ABB RAPID module: MainProgram.mod

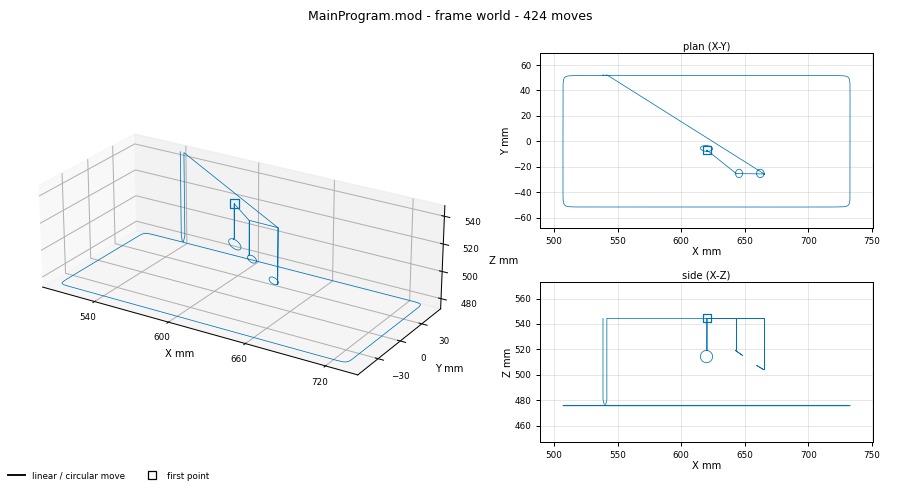
[picture p0: tool path of MainProgram.mod in frame world, 424 of 456 moves have a stored position in this frame; points joined in program order, loops and branches not executed]
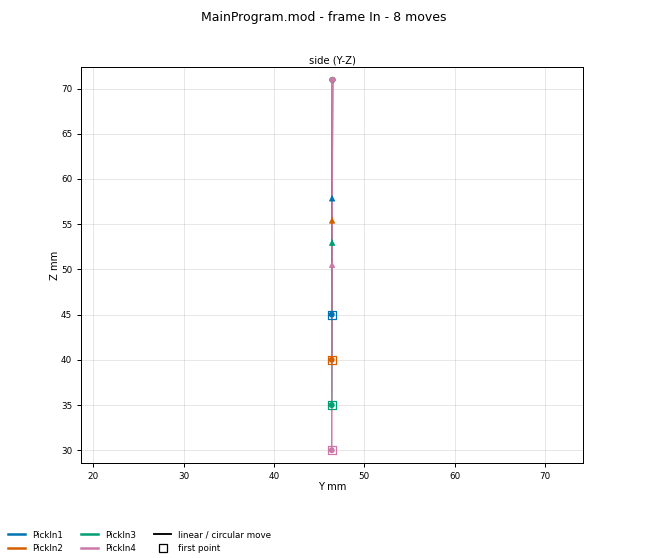
[picture p1: tool path of MainProgram.mod in frame In, 8 of 456 moves have a stored position in this frame; points joined in program order, loops and branches not executed]
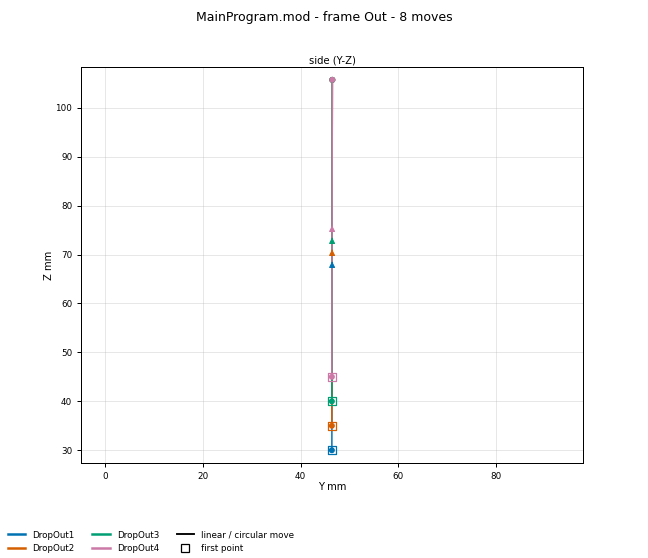
[picture p2: tool path of MainProgram.mod in frame Out, 8 of 456 moves have a stored position in this frame; points joined in program order, loops and branches not executed]
%%%
  VERSION:1
  LANGUAGE:ENGLISH
%%%
MODULE MOD_MainProgram

    ! -------------------------------
    ! Define customized variables here
    ! ...

	! Tool variables:
	PERS tooldata SuctionCup := [TRUE,[[-94.709,0.000,259.352],[0.00000000,0.00000000,0.00000000,1.00000000]],[1,[0,0,20],[1,0,0,0],0,0,0.005]];
	PERS tooldata Spindle := [TRUE,[[186.140,-0.004,258.607],[0.87136628,0.00000000,0.49063307,0.00000000]],[1,[0,0,20],[1,0,0,0],0,0,0.005]];

	! Reference variables:
	PERS wobjdata World := [FALSE, TRUE, "", [[0,0,0],[1,0,0,0]],[[390.000,0.000,0.000],[1.00000000,0.00000000,0.00000000,0.00000000]]];
	PERS wobjdata In := [FALSE, TRUE, "", [[0,0,0],[1,0,0,0]],[[290.000,450.000,10.000],[1.00000000,0.00000000,0.00000000,0.00000000]]];
	PERS wobjdata PartStation := [FALSE, TRUE, "", [[0,0,0],[1,0,0,0]],[[620.000,0.000,396.884],[0.70710678,0.00000000,0.00000000,-0.70710678]]];
	PERS wobjdata Deburring := [FALSE, TRUE, "", [[0,0,0],[1,0,0,0]],[[620.000,0.000,458.384],[0.70710678,0.00000000,0.00000000,-0.70710678]]];
	PERS wobjdata Out := [FALSE, TRUE, "", [[0,0,0],[1,0,0,0]],[[290.000,-450.000,10.000],[1.00000000,0.00000000,0.00000000,0.00000000]]];

	PROC GoHome()
		ConfJ \On;
		ConfL \Off;
		World := [FALSE, TRUE, "", [[0,0,0],[1,0,0,0]],[[390.000,0.000,0.000],[1.00000000,0.00000000,0.00000000,0.00000000]]];
		MoveAbsJ [[0.000000,0.000000,-20.000000,0.000000,30.170000,0.000000],[9E+09,9E+09,9E+09,9E+09,9E+09,9E+09]],v500,z1,SuctionCup \WObj:=World;
	ENDPROC

	PROC PickIn1()
		ConfJ \On;
		ConfL \Off;
		SuctionCup := [TRUE,[[-94.709,0.000,259.352],[0.00000000,0.00000000,0.00000000,1.00000000]],[1,[0,0,20],[1,0,0,0],0,0,0.005]];
		MoveAbsJ [[70.152800,32.938500,23.515600,0.000000,33.545900,70.152800],[9E+09,9E+09,9E+09,9E+09,9E+09,9E+09]],v500,z1,SuctionCup \WObj:=In;
		MoveL [[-16.111,46.392,45.000],[0.00000000,1.00000000,0.00000000,-0.00000000],[0,2,-2,1],[9E+09,9E+09,9E+09,9E+09,9E+09,9E+09]],v500,z1,SuctionCup \WObj:=In;
		! Attach to Suction Cup
		WaitTime 0.500;
		MoveL [[-16.087,46.472,70.960],[0.00000000,1.00000000,0.00000000,-0.00000000],[0,0,0,0],[9E+09,9E+09,9E+09,9E+09,9E+09,9E+09]],v500,z1,SuctionCup \WObj:=In;
	ENDPROC

	PROC DropStation()
		ConfJ \On;
		ConfL \Off;
		SuctionCup := [TRUE,[[-94.709,0.000,259.352],[0.00000000,0.00000000,0.00000000,1.00000000]],[1,[0,0,20],[1,0,0,0],0,0,0.005]];
		MoveAbsJ [[9.440500,34.191600,-49.511700,0.000000,105.320000,99.440500],[9E+09,9E+09,9E+09,9E+09,9E+09,9E+09]],v500,z1,SuctionCup \WObj:=PartStation;
		MoveL [[-16.111,46.392,100.500],[0.00000000,1.00000000,0.00000000,-0.00000000],[0,2,-1,1],[9E+09,9E+09,9E+09,9E+09,9E+09,9E+09]],v500,z1,SuctionCup \WObj:=PartStation;
		! Detach from Suction Cup
		WaitTime 0.500;
		MoveL [[-16.111,46.485,191.000],[0.00000000,1.00000000,0.00000000,-0.00000000],[0,0,1,0],[9E+09,9E+09,9E+09,9E+09,9E+09,9E+09]],v500,z1,SuctionCup \WObj:=PartStation;
	ENDPROC

	PROC Station1()
		ConfJ \On;
		ConfL \Off;
		! show Spindle
		TPWrite "/'Plastic deburring v9'";
		TPWrite "/''";
		TPWrite "/'NEW SECTION'";
		TPWrite "/'Strategy: swarf5d'";
		TPWrite "/'Comment: Swarf8'";
		TPWrite "/'MATRIX DEFINITION'";
		TPWrite "/'Output x(i),y(i),z(i)'";
		TPWrite "/'Output x(j),y(j),z(j)'";
		TPWrite "/'Output x(k),y(k),z(k)'";
		TPWrite "/'Output dx,dy,dz'";
		SetTool 3;
		SetRPM 5000.0;
		Spindle 1;
		MoveAbsJ [[35.301800,13.650800,12.157300,-89.295200,63.027800,42.556000],[9E+09,9E+09,9E+09,9E+09,9E+09,9E+09]],v1000,z1,Spindle \WObj:=Deburring;
		MoveL [[6.917,0.414,86.000],[0.38548738,-0.58483375,0.59278955,-0.39745378],[0,-1,0,0],[9E+09,9E+09,9E+09,9E+09,9E+09,9E+09]],v1000,z1,Spindle \WObj:=Deburring;
		MoveL [[6.917,0.414,86.000],[0.38548738,-0.58483375,0.59278955,-0.39745378],[0,-1,0,0],[9E+09,9E+09,9E+09,9E+09,9E+09,9E+09]],v1000,z1,Spindle \WObj:=Deburring;
		MoveL [[6.917,0.414,61.098],[0.38548738,-0.58483375,0.59278955,-0.39745378],[0,-2,0,0],[9E+09,9E+09,9E+09,9E+09,9E+09,9E+09]],v1000,z1,Spindle \WObj:=Deburring;
		MoveL [[7.874,0.393,60.697],[0.38548738,-0.58483375,0.59278955,-0.39745378],[0,-2,0,0],[9E+09,9E+09,9E+09,9E+09,9E+09,9E+09]],[16.67,500,5000,1000],z1,Spindle \WObj:=Deburring;
		MoveL [[7.903,0.385,60.695],[0.38548738,-0.58483375,0.59278955,-0.39745378],[0,-2,0,0],[9E+09,9E+09,9E+09,9E+09,9E+09,9E+09]],[16.67,500,5000,1000],z1,Spindle \WObj:=Deburring;
		MoveL [[7.923,0.368,60.712],[0.38548738,-0.58483375,0.59278955,-0.39745378],[0,-2,0,0],[9E+09,9E+09,9E+09,9E+09,9E+09,9E+09]],[16.67,500,5000,1000],z1,Spindle \WObj:=Deburring;
		MoveL [[7.932,0.350,60.736],[0.38548738,-0.58483375,0.59278955,-0.39745378],[0,-2,0,0],[9E+09,9E+09,9E+09,9E+09,9E+09,9E+09]],[16.67,500,5000,1000],z1,Spindle \WObj:=Deburring;
		MoveL [[7.942,0.339,60.763],[0.38548738,-0.58483375,0.59278955,-0.39745378],[0,-2,0,0],[9E+09,9E+09,9E+09,9E+09,9E+09,9E+09]],[16.67,500,5000,1000],z1,Spindle \WObj:=Deburring;
		MoveL [[7.946,0.311,60.775],[0.38548738,-0.58483375,0.59278955,-0.39745378],[0,-2,0,0],[9E+09,9E+09,9E+09,9E+09,9E+09,9E+09]],[16.67,500,5000,1000],z1,Spindle \WObj:=Deburring;
		MoveL [[7.938,0.025,60.788],[0.38288630,-0.58214828,0.59447297,-0.40137683],[0,-2,0,0],[9E+09,9E+09,9E+09,9E+09,9E+09,9E+09]],[16.67,500,5000,1000],z1,Spindle \WObj:=Deburring;
		MoveL [[7.910,-0.405,60.779],[0.38300483,-0.58012093,0.59439635,-0.40430185],[0,-2,0,0],[9E+09,9E+09,9E+09,9E+09,9E+09,9E+09]],[16.67,500,5000,1000],z1,Spindle \WObj:=Deburring;
		MoveL [[7.848,-0.934,60.707],[0.38194021,-0.57666146,0.59508111,-0.40922086],[0,-2,0,0],[9E+09,9E+09,9E+09,9E+09,9E+09,9E+09]],[16.67,500,5000,1000],z1,Spindle \WObj:=Deburring;
		MoveL [[7.772,-1.372,60.601],[0.37995322,-0.57413190,0.59635187,-0.41276211],[0,-1,0,0],[9E+09,9E+09,9E+09,9E+09,9E+09,9E+09]],[16.67,500,5000,1000],z1,Spindle \WObj:=Deburring;
		MoveL [[7.660,-1.869,60.426],[0.37743363,-0.57188089,0.59794992,-0.41587499],[0,-1,0,0],[9E+09,9E+09,9E+09,9E+09,9E+09,9E+09]],[16.67,500,5000,1000],z1,Spindle \WObj:=Deburring;
		MoveL [[7.526,-2.338,60.200],[0.37439771,-0.57017304,0.59985541,-0.41821351],[0,-1,0,0],[9E+09,9E+09,9E+09,9E+09,9E+09,9E+09]],[16.67,500,5000,1000],z1,Spindle \WObj:=Deburring;
		MoveL [[7.336,-2.857,59.865],[0.36917090,-0.56926904,0.60308585,-0.41944375],[0,-1,0,0],[9E+09,9E+09,9E+09,9E+09,9E+09,9E+09]],[16.67,500,5000,1000],z1,Spindle \WObj:=Deburring;
		MoveL [[7.162,-3.251,59.544],[0.36551673,-0.56883653,0.60530778,-0.42002978],[0,-1,0,0],[9E+09,9E+09,9E+09,9E+09,9E+09,9E+09]],[16.67,500,5000,1000],z1,Spindle \WObj:=Deburring;
		MoveL [[6.973,-3.606,59.186],[0.36224838,-0.56788024,0.60726923,-0.42132199],[0,-1,0,0],[9E+09,9E+09,9E+09,9E+09,9E+09,9E+09]],[16.67,500,5000,1000],z1,Spindle \WObj:=Deburring;
		MoveL [[6.815,-3.864,58.879],[0.36043999,-0.56727725,0.60834425,-0.42213363],[0,-1,0,0],[9E+09,9E+09,9E+09,9E+09,9E+09,9E+09]],[16.67,500,5000,1000],z1,Spindle \WObj:=Deburring;
		MoveL [[6.554,-4.204,58.361],[0.35672537,-0.56741746,0.61052971,-0.42194538],[0,-1,0,0],[9E+09,9E+09,9E+09,9E+09,9E+09,9E+09]],[16.67,500,5000,1000],z1,Spindle \WObj:=Deburring;
		MoveL [[6.282,-4.474,57.808],[0.35340770,-0.56800021,0.61245687,-0.42115952],[0,-1,0,0],[9E+09,9E+09,9E+09,9E+09,9E+09,9E+09]],[16.67,500,5000,1000],z1,Spindle \WObj:=Deburring;
		MoveL [[6.084,-4.622,57.400],[0.35045021,-0.56898176,0.61415334,-0.41983338],[0,-1,0,0],[9E+09,9E+09,9E+09,9E+09,9E+09,9E+09]],[16.67,500,5000,1000],z1,Spindle \WObj:=Deburring;
		MoveL [[5.801,-4.764,56.806],[0.34689032,-0.56972554,0.61617155,-0.41882280],[0,-1,0,0],[9E+09,9E+09,9E+09,9E+09,9E+09,9E+09]],[16.67,500,5000,1000],z1,Spindle \WObj:=Deburring;
		MoveL [[5.517,-4.832,56.200],[0.34354127,-0.57095868,0.61804469,-0.41714067],[0,-1,0,0],[9E+09,9E+09,9E+09,9E+09,9E+09,9E+09]],[16.67,500,5000,1000],z1,Spindle \WObj:=Deburring;
		MoveL [[5.234,-4.822,55.590],[0.34057760,-0.57257464,0.61968277,-0.41491981],[0,-1,0,0],[9E+09,9E+09,9E+09,9E+09,9E+09,9E+09]],[16.67,500,5000,1000],z1,Spindle \WObj:=Deburring;
		MoveL [[4.956,-4.736,54.983],[0.33797772,-0.57446132,0.62110430,-0.41230413],[0,-1,0,0],[9E+09,9E+09,9E+09,9E+09,9E+09,9E+09]],[16.67,500,5000,1000],z1,Spindle \WObj:=Deburring;
		MoveL [[4.687,-4.572,54.389],[0.33604086,-0.57652798,0.62215522,-0.40940801],[0,-1,0,0],[9E+09,9E+09,9E+09,9E+09,9E+09,9E+09]],[16.67,500,5000,1000],z1,Spindle \WObj:=Deburring;
		MoveL [[4.440,-4.339,53.840],[0.33425295,-0.57979674,0.62311733,-0.40476598],[0,-1,0,0],[9E+09,9E+09,9E+09,9E+09,9E+09,9E+09]],[16.67,500,5000,1000],z1,Spindle \WObj:=Deburring;
		MoveL [[4.245,-4.095,53.402],[0.33283353,-0.58190363,0.62387648,-0.40173143],[0,-1,0,0],[9E+09,9E+09,9E+09,9E+09,9E+09,9E+09]],[16.67,500,5000,1000],z1,Spindle \WObj:=Deburring;
		MoveL [[4.097,-3.868,53.067],[0.33181431,-0.58289839,0.62441871,-0.40028740],[0,-1,0,0],[9E+09,9E+09,9E+09,9E+09,9E+09,9E+09]],[16.67,500,5000,1000],z1,Spindle \WObj:=Deburring;
		MoveL [[3.907,-3.500,52.631],[0.32892812,-0.58510481,0.62594413,-0.39705490],[0,-1,0,0],[9E+09,9E+09,9E+09,9E+09,9E+09,9E+09]],[16.67,500,5000,1000],z1,Spindle \WObj:=Deburring;
		MoveL [[3.755,-3.123,52.278],[0.32712779,-0.58752921,0.62688678,-0.39345876],[0,-1,0,0],[9E+09,9E+09,9E+09,9E+09,9E+09,9E+09]],[16.67,500,5000,1000],z1,Spindle \WObj:=Deburring;
		MoveL [[3.623,-2.706,51.964],[0.32579005,-0.59003824,0.62758358,-0.38968521],[0,-1,0,0],[9E+09,9E+09,9E+09,9E+09,9E+09,9E+09]],[16.67,500,5000,1000],z1,Spindle \WObj:=Deburring;
		MoveL [[3.513,-2.253,51.695],[0.32545472,-0.59261817,0.62775754,-0.38575044],[0,-1,0,0],[9E+09,9E+09,9E+09,9E+09,9E+09,9E+09]],[16.67,500,5000,1000],z1,Spindle \WObj:=Deburring;
		MoveL [[3.426,-1.769,51.476],[0.32546867,-0.59528891,0.62774999,-0.38161657],[0,-1,0,0],[9E+09,9E+09,9E+09,9E+09,9E+09,9E+09]],[16.67,500,5000,1000],z1,Spindle \WObj:=Deburring;
		MoveL [[3.367,-1.261,51.311],[0.32642133,-0.59790109,0.62725498,-0.37751104],[0,-1,0,0],[9E+09,9E+09,9E+09,9E+09,9E+09,9E+09]],[16.67,500,5000,1000],z1,Spindle \WObj:=Deburring;
		MoveL [[3.336,-0.734,51.202],[0.32721447,-0.60077200,0.62684183,-0.37292496],[0,-1,0,0],[9E+09,9E+09,9E+09,9E+09,9E+09,9E+09]],[16.67,500,5000,1000],z1,Spindle \WObj:=Deburring;
		MoveL [[3.334,-0.198,51.154],[0.32817251,-0.60371090,0.62634061,-0.36814859],[0,-1,0,0],[9E+09,9E+09,9E+09,9E+09,9E+09,9E+09]],[16.67,500,5000,1000],z1,Spindle \WObj:=Deburring;
		MoveL [[3.362,0.339,51.167],[0.32965343,-0.60642410,0.62556274,-0.36366150],[0,-1,0,0],[9E+09,9E+09,9E+09,9E+09,9E+09,9E+09]],[16.67,500,5000,1000],z1,Spindle \WObj:=Deburring;
		MoveL [[3.419,0.869,51.239],[0.33178536,-0.60854381,0.62443456,-0.36010330],[0,-1,0,0],[9E+09,9E+09,9E+09,9E+09,9E+09,9E+09]],[16.67,500,5000,1000],z1,Spindle \WObj:=Deburring;
		MoveL [[3.511,1.417,51.385],[0.33673317,-0.61021010,0.62178053,-0.35727213],[0,-1,0,0],[9E+09,9E+09,9E+09,9E+09,9E+09,9E+09]],[16.67,500,5000,1000],z1,Spindle \WObj:=Deburring;
		MoveL [[3.596,1.815,51.527],[0.33843795,-0.61063438,0.62085393,-0.35654705],[0,-1,0,0],[9E+09,9E+09,9E+09,9E+09,9E+09,9E+09]],[16.67,500,5000,1000],z1,Spindle \WObj:=Deburring;
		MoveL [[3.725,2.284,51.756],[0.34227325,-0.61131950,0.61874797,-0.35537084],[0,-1,0,0],[9E+09,9E+09,9E+09,9E+09,9E+09,9E+09]],[16.67,500,5000,1000],z1,Spindle \WObj:=Deburring;
		MoveL [[3.876,2.722,52.031],[0.34580120,-0.61257678,0.61678310,-0.35319942],[0,-1,0,0],[9E+09,9E+09,9E+09,9E+09,9E+09,9E+09]],[16.67,500,5000,1000],z1,Spindle \WObj:=Deburring;
		MoveL [[4.045,3.123,52.347],[0.34927682,-0.61344264,0.61482152,-0.35169353],[0,-1,0,0],[9E+09,9E+09,9E+09,9E+09,9E+09,9E+09]],[16.67,500,5000,1000],z1,Spindle \WObj:=Deburring;
		MoveL [[4.270,3.549,52.777],[0.35456914,-0.61410907,0.61178476,-0.35052844],[0,-1,0,0],[9E+09,9E+09,9E+09,9E+09,9E+09,9E+09]],[16.67,500,5000,1000],z1,Spindle \WObj:=Deburring;
		MoveL [[4.470,3.860,53.168],[0.35787236,-0.61441666,0.60985864,-0.34998855],[0,-1,0,0],[9E+09,9E+09,9E+09,9E+09,9E+09,9E+09]],[16.67,500,5000,1000],z1,Spindle \WObj:=Deburring;
		MoveL [[4.682,4.127,53.589],[0.36134434,-0.61410206,0.60780784,-0.35054039],[0,-1,0,0],[9E+09,9E+09,9E+09,9E+09,9E+09,9E+09]],[16.67,500,5000,1000],z1,Spindle \WObj:=Deburring;
		MoveL [[4.909,4.360,54.045],[0.36290006,-0.61402146,0.60688026,-0.35068155],[0,-1,0,0],[9E+09,9E+09,9E+09,9E+09,9E+09,9E+09]],[16.67,500,5000,1000],z1,Spindle \WObj:=Deburring;
		MoveL [[5.207,4.574,54.652],[0.36756237,-0.61295146,0.60406786,-0.35254849],[0,-2,0,0],[9E+09,9E+09,9E+09,9E+09,9E+09,9E+09]],[16.67,500,5000,1000],z1,Spindle \WObj:=Deburring;
		MoveL [[5.440,4.682,55.130],[0.37069589,-0.61194017,0.60215000,-0.35430095],[0,-2,0,0],[9E+09,9E+09,9E+09,9E+09,9E+09,9E+09]],[16.67,500,5000,1000],z1,Spindle \WObj:=Deburring;
		MoveL [[5.682,4.750,55.631],[0.37301034,-0.61212853,0.60071915,-0.35397521],[0,-2,0,0],[9E+09,9E+09,9E+09,9E+09,9E+09,9E+09]],[16.67,500,5000,1000],z1,Spindle \WObj:=Deburring;
		MoveL [[5.972,4.756,56.238],[0.37688431,-0.61142117,0.59829589,-0.35519628],[0,-2,0,0],[9E+09,9E+09,9E+09,9E+09,9E+09,9E+09]],[16.67,500,5000,1000],z1,Spindle \WObj:=Deburring;
		MoveL [[6.258,4.684,56.843],[0.38040882,-0.61035480,0.59606153,-0.35702493],[0,-2,0,0],[9E+09,9E+09,9E+09,9E+09,9E+09,9E+09]],[16.67,500,5000,1000],z1,Spindle \WObj:=Deburring;
		MoveL [[6.536,4.537,57.438],[0.38298801,-0.60875341,0.59440720,-0.35974929],[0,-2,0,0],[9E+09,9E+09,9E+09,9E+09,9E+09,9E+09]],[16.67,500,5000,1000],z1,Spindle \WObj:=Deburring;
		MoveL [[6.802,4.313,58.013],[0.38480474,-0.60692696,0.59323291,-0.36282185],[0,-2,0,0],[9E+09,9E+09,9E+09,9E+09,9E+09,9E+09]],[16.67,500,5000,1000],z1,Spindle \WObj:=Deburring;
		MoveL [[7.042,4.024,58.538],[0.38647889,-0.60399208,0.59214367,-0.36768670],[0,-2,0,0],[9E+09,9E+09,9E+09,9E+09,9E+09,9E+09]],[16.67,500,5000,1000],z1,Spindle \WObj:=Deburring;
		MoveL [[7.193,3.799,58.873],[0.38664149,-0.60298907,0.59203745,-0.36932938],[0,-2,0,0],[9E+09,9E+09,9E+09,9E+09,9E+09,9E+09]],[16.67,500,5000,1000],z1,Spindle \WObj:=Deburring;
		MoveL [[7.386,3.431,59.308],[0.38767021,-0.60080000,0.59136449,-0.37287962],[0,-2,0,0],[9E+09,9E+09,9E+09,9E+09,9E+09,9E+09]],[16.67,500,5000,1000],z1,Spindle \WObj:=Deburring;
		MoveL [[7.541,3.055,59.661],[0.38899214,-0.59839293,0.59049568,-0.37673051],[0,-2,0,0],[9E+09,9E+09,9E+09,9E+09,9E+09,9E+09]],[16.67,500,5000,1000],z1,Spindle \WObj:=Deburring;
		MoveL [[7.675,2.640,59.976],[0.39067221,-0.59591183,0.58938556,-0.38064284],[0,-2,0,0],[9E+09,9E+09,9E+09,9E+09,9E+09,9E+09]],[16.67,500,5000,1000],z1,Spindle \WObj:=Deburring;
		MoveL [[7.785,2.187,60.246],[0.39103498,-0.59339095,0.58914492,-0.38456089],[0,-2,0,0],[9E+09,9E+09,9E+09,9E+09,9E+09,9E+09]],[16.67,500,5000,1000],z1,Spindle \WObj:=Deburring;
		MoveL [[7.869,1.704,60.467],[0.39061269,-0.59084673,0.58942483,-0.38845881],[0,-2,0,0],[9E+09,9E+09,9E+09,9E+09,9E+09,9E+09]],[16.67,500,5000,1000],z1,Spindle \WObj:=Deburring;
		MoveL [[7.924,1.195,60.633],[0.38860975,-0.58858373,0.59074741,-0.39187901],[0,-2,0,0],[9E+09,9E+09,9E+09,9E+09,9E+09,9E+09]],[16.67,500,5000,1000],z1,Spindle \WObj:=Deburring;
		MoveL [[7.949,0.668,60.742],[0.38626315,-0.58624691,0.59228428,-0.39536650],[0,-2,0,0],[9E+09,9E+09,9E+09,9E+09,9E+09,9E+09]],[16.67,500,5000,1000],z1,Spindle \WObj:=Deburring;
		MoveL [[7.948,0.549,60.753],[0.38498996,-0.58493913,0.59311268,-0.39729875],[0,-2,0,0],[9E+09,9E+09,9E+09,9E+09,9E+09,9E+09]],[16.67,500,5000,1000],z1,Spindle \WObj:=Deburring;
		MoveL [[7.947,0.430,60.764],[0.38524128,-0.58488478,0.59294941,-0.39737884],[0,-2,0,0],[9E+09,9E+09,9E+09,9E+09,9E+09,9E+09]],[16.67,500,5000,1000],z1,Spindle \WObj:=Deburring;
		MoveL [[7.946,0.311,60.775],[0.38548738,-0.58483375,0.59278955,-0.39745378],[0,-2,0,0],[9E+09,9E+09,9E+09,9E+09,9E+09,9E+09]],[16.67,500,5000,1000],z1,Spindle \WObj:=Deburring;
		MoveL [[7.941,0.282,60.765],[0.38548738,-0.58483375,0.59278955,-0.39745378],[0,-2,0,0],[9E+09,9E+09,9E+09,9E+09,9E+09,9E+09]],[16.67,500,5000,1000],z1,Spindle \WObj:=Deburring;
		MoveL [[7.929,0.270,60.740],[0.38548738,-0.58483375,0.59278955,-0.39745378],[0,-2,0,0],[9E+09,9E+09,9E+09,9E+09,9E+09,9E+09]],[16.67,500,5000,1000],z1,Spindle \WObj:=Deburring;
		MoveL [[7.919,0.250,60.718],[0.38548738,-0.58483375,0.59278955,-0.39745378],[0,-2,0,0],[9E+09,9E+09,9E+09,9E+09,9E+09,9E+09]],[16.67,500,5000,1000],z1,Spindle \WObj:=Deburring;
		MoveL [[7.900,0.232,60.703],[0.38548738,-0.58483375,0.59278955,-0.39745378],[0,-2,0,0],[9E+09,9E+09,9E+09,9E+09,9E+09,9E+09]],[16.67,500,5000,1000],z1,Spindle \WObj:=Deburring;
		MoveL [[7.870,0.225,60.706],[0.38548738,-0.58483375,0.59278955,-0.39745378],[0,-2,0,0],[9E+09,9E+09,9E+09,9E+09,9E+09,9E+09]],[16.67,500,5000,1000],z1,Spindle \WObj:=Deburring;
		MoveL [[7.870,0.225,60.706],[0.38548738,-0.58483375,0.59278955,-0.39745378],[0,-2,0,0],[9E+09,9E+09,9E+09,9E+09,9E+09,9E+09]],v1000,z1,Spindle \WObj:=Deburring;
		MoveL [[6.903,0.247,61.111],[0.38548738,-0.58483375,0.59278955,-0.39745378],[0,-2,0,0],[9E+09,9E+09,9E+09,9E+09,9E+09,9E+09]],v1000,z1,Spindle \WObj:=Deburring;
		MoveL [[6.903,0.247,86.000],[0.38548738,-0.58483375,0.59278955,-0.39745378],[0,-1,0,0],[9E+09,9E+09,9E+09,9E+09,9E+09,9E+09]],v1000,z1,Spindle \WObj:=Deburring;
		TPWrite "/'NEW SECTION'";
		TPWrite "/'Strategy: swarf5d'";
		TPWrite "/'Comment: Swarf9'";
		TPWrite "/'MATRIX DEFINITION'";
		TPWrite "/'Output x(i),y(i),z(i)'";
		TPWrite "/'Output x(j),y(j),z(j)'";
		TPWrite "/'Output x(k),y(k),z(k)'";
		TPWrite "/'Output dx,dy,dz'";
		SetTool 3;
		SetRPM 5000.0;
		MoveL [[25.588,23.564,86.000],[0.22593931,0.66585901,-0.67003984,0.23797020],[-1,-1,-1,0],[9E+09,9E+09,9E+09,9E+09,9E+09,9E+09]],v1000,z1,Spindle \WObj:=Deburring;
		MoveL [[25.588,23.564,61.477],[0.22593931,0.66585901,-0.67003984,0.23797020],[-1,-1,-1,0],[9E+09,9E+09,9E+09,9E+09,9E+09,9E+09]],v1000,z1,Spindle \WObj:=Deburring;
		MoveL [[25.602,22.924,60.668],[0.22593931,0.66585901,-0.67003984,0.23797020],[-1,-1,-1,0],[9E+09,9E+09,9E+09,9E+09,9E+09,9E+09]],[16.67,500,5000,1000],z1,Spindle \WObj:=Deburring;
		MoveL [[25.596,22.899,60.651],[0.22593931,0.66585901,-0.67003984,0.23797020],[-1,-1,-1,0],[9E+09,9E+09,9E+09,9E+09,9E+09,9E+09]],[16.67,500,5000,1000],z1,Spindle \WObj:=Deburring;
		MoveL [[25.580,22.874,60.656],[0.22593931,0.66585901,-0.67003984,0.23797020],[-1,-1,-1,0],[9E+09,9E+09,9E+09,9E+09,9E+09,9E+09]],[16.67,500,5000,1000],z1,Spindle \WObj:=Deburring;
		MoveL [[25.561,22.854,60.672],[0.22593931,0.66585901,-0.67003984,0.23797020],[-1,-1,-1,0],[9E+09,9E+09,9E+09,9E+09,9E+09,9E+09]],[16.67,500,5000,1000],z1,Spindle \WObj:=Deburring;
		MoveL [[25.551,22.831,60.690],[0.22593931,0.66585901,-0.67003984,0.23797020],[-1,-1,-1,0],[9E+09,9E+09,9E+09,9E+09,9E+09,9E+09]],[16.67,500,5000,1000],z1,Spindle \WObj:=Deburring;
		MoveL [[25.523,22.821,60.698],[0.22593931,0.66585901,-0.67003984,0.23797020],[-1,-1,-1,0],[9E+09,9E+09,9E+09,9E+09,9E+09,9E+09]],[16.67,500,5000,1000],z1,Spindle \WObj:=Deburring;
		MoveL [[25.288,22.812,60.703],[0.23132418,0.66725233,-0.66819988,0.23403496],[-1,0,-1,0],[9E+09,9E+09,9E+09,9E+09,9E+09,9E+09]],[16.67,500,5000,1000],z1,Spindle \WObj:=Deburring;
		MoveL [[24.985,22.820,60.698],[0.23450445,0.66763618,-0.66709034,0.23293793],[-1,0,-1,0],[9E+09,9E+09,9E+09,9E+09,9E+09,9E+09]],[16.67,500,5000,1000],z1,Spindle \WObj:=Deburring;
		MoveL [[24.587,22.871,60.663],[0.24007837,0.66885645,-0.66510328,0.22941457],[-1,0,-1,0],[9E+09,9E+09,9E+09,9E+09,9E+09,9E+09]],[16.67,500,5000,1000],z1,Spindle \WObj:=Deburring;
		MoveL [[24.199,22.964,60.601],[0.24468394,0.67027520,-0.66342218,0.22523751],[-1,0,-1,0],[9E+09,9E+09,9E+09,9E+09,9E+09,9E+09]],[16.67,500,5000,1000],z1,Spindle \WObj:=Deburring;
		MoveL [[23.827,23.095,60.514],[0.24823939,0.67184973,-0.66209949,0.22049811],[-1,0,-1,0],[9E+09,9E+09,9E+09,9E+09,9E+09,9E+09]],[16.67,500,5000,1000],z1,Spindle \WObj:=Deburring;
		MoveL [[23.397,23.314,60.369],[0.25136263,0.67436154,-0.66092270,0.21268411],[-1,0,-1,0],[9E+09,9E+09,9E+09,9E+09,9E+09,9E+09]],[16.67,500,5000,1000],z1,Spindle \WObj:=Deburring;
		MoveL [[23.082,23.524,60.229],[0.25221713,0.67605558,-0.66059650,0.20723812],[-1,0,-1,0],[9E+09,9E+09,9E+09,9E+09,9E+09,9E+09]],[16.67,500,5000,1000],z1,Spindle \WObj:=Deburring;
		MoveL [[22.801,23.764,60.067],[0.25279268,0.67777283,-0.66037454,0.20155723],[-1,0,-1,0],[9E+09,9E+09,9E+09,9E+09,9E+09,9E+09]],[16.67,500,5000,1000],z1,Spindle \WObj:=Deburring;
		MoveL [[22.556,24.029,59.887],[0.25451140,0.67948076,-0.65971680,0.19571305],[-1,0,-1,0],[9E+09,9E+09,9E+09,9E+09,9E+09,9E+09]],[16.67,500,5000,1000],z1,Spindle \WObj:=Deburring;
		MoveL [[22.351,24.316,59.691],[0.25639160,0.68117668,-0.65898852,0.18972564],[-1,0,-1,0],[9E+09,9E+09,9E+09,9E+09,9E+09,9E+09]],[16.67,500,5000,1000],z1,Spindle \WObj:=Deburring;
		MoveL [[22.188,24.620,59.482],[0.25707629,0.68268733,-0.65871885,0.18422614],[-1,0,-1,0],[9E+09,9E+09,9E+09,9E+09,9E+09,9E+09]],[16.67,500,5000,1000],z1,Spindle \WObj:=Deburring;
		MoveL [[22.070,24.937,59.263],[0.25603932,0.68390940,-0.65912393,0.17963142],[-1,0,-1,0],[9E+09,9E+09,9E+09,9E+09,9E+09,9E+09]],[16.67,500,5000,1000],z1,Spindle \WObj:=Deburring;
		MoveL [[21.999,25.263,59.037],[0.25372125,0.68489416,-0.66001913,0.17584158],[-1,0,-1,0],[9E+09,9E+09,9E+09,9E+09,9E+09,9E+09]],[16.67,500,5000,1000],z1,Spindle \WObj:=Deburring;
		MoveL [[21.974,25.593,58.807],[0.25059987,0.68561674,-0.66121165,0.17299871],[-1,0,-1,0],[9E+09,9E+09,9E+09,9E+09,9E+09,9E+09]],[16.67,500,5000,1000],z1,Spindle \WObj:=Deburring;
		MoveL [[21.997,25.924,58.577],[0.24620099,0.68599910,-0.66286170,0.17147791],[-1,0,-1,0],[9E+09,9E+09,9E+09,9E+09,9E+09,9E+09]],[16.67,500,5000,1000],z1,Spindle \WObj:=Deburring;
		MoveL [[22.067,26.248,58.349],[0.24109769,0.68616380,-0.66473597,0.17081344],[-1,0,-1,0],[9E+09,9E+09,9E+09,9E+09,9E+09,9E+09]],[16.67,500,5000,1000],z1,Spindle \WObj:=Deburring;
		MoveL [[22.184,26.564,58.126],[0.23603372,0.68628710,-0.66655055,0.17031872],[-1,0,-1,0],[9E+09,9E+09,9E+09,9E+09,9E+09,9E+09]],[16.67,500,5000,1000],z1,Spindle \WObj:=Deburring;
		MoveL [[22.345,26.865,57.913],[0.23111847,0.68648459,-0.66826955,0.16952572],[-1,0,-1,0],[9E+09,9E+09,9E+09,9E+09,9E+09,9E+09]],[16.67,500,5000,1000],z1,Spindle \WObj:=Deburring;
		MoveL [[22.549,27.149,57.711],[0.22656366,0.68660155,-0.66982723,0.16905237],[-1,0,-1,0],[9E+09,9E+09,9E+09,9E+09,9E+09,9E+09]],[16.67,500,5000,1000],z1,Spindle \WObj:=Deburring;
		MoveL [[22.608,27.216,57.663],[0.22665394,0.68656149,-0.66979846,0.16920796],[-1,0,-1,0],[9E+09,9E+09,9E+09,9E+09,9E+09,9E+09]],[16.67,500,5000,1000],z1,Spindle \WObj:=Deburring;
		MoveL [[22.666,27.282,57.615],[0.22673822,0.68652339,-0.66976819,0.16936938],[-1,0,-1,0],[9E+09,9E+09,9E+09,9E+09,9E+09,9E+09]],[16.67,500,5000,1000],z1,Spindle \WObj:=Deburring;
		MoveL [[22.725,27.349,57.568],[0.22391864,0.68648721,-0.67071733,0.16951112],[-1,0,-1,0],[9E+09,9E+09,9E+09,9E+09,9E+09,9E+09]],[16.67,500,5000,1000],z1,Spindle \WObj:=Deburring;
		MoveL [[23.076,27.643,57.356],[0.21586440,0.68640623,-0.67335239,0.16983994],[-1,0,-1,0],[9E+09,9E+09,9E+09,9E+09,9E+09,9E+09]],[16.67,500,5000,1000],z1,Spindle \WObj:=Deburring;
		MoveL [[23.390,27.848,57.209],[0.21073883,0.68641279,-0.67497178,0.16982263],[-1,0,-1,0],[9E+09,9E+09,9E+09,9E+09,9E+09,9E+09]],[16.67,500,5000,1000],z1,Spindle \WObj:=Deburring;
		MoveL [[23.733,28.021,57.084],[0.20571489,0.68624503,-0.67652291,0.17048721],[-1,0,-1,0],[9E+09,9E+09,9E+09,9E+09,9E+09,9E+09]],[16.67,500,5000,1000],z1,Spindle \WObj:=Deburring;
		MoveL [[24.099,28.158,56.986],[0.20112152,0.68565538,-0.67790262,0.17284351],[-1,0,-1,0],[9E+09,9E+09,9E+09,9E+09,9E+09,9E+09]],[16.67,500,5000,1000],z1,Spindle \WObj:=Deburring;
		MoveL [[24.483,28.257,56.914],[0.19703903,0.68466952,-0.67909945,0.17671224],[-1,0,-1,0],[9E+09,9E+09,9E+09,9E+09,9E+09,9E+09]],[16.67,500,5000,1000],z1,Spindle \WObj:=Deburring;
		MoveL [[24.879,28.318,56.871],[0.19320632,0.68349149,-0.68020030,0.18121325],[-1,0,-1,0],[9E+09,9E+09,9E+09,9E+09,9E+09,9E+09]],[16.67,500,5000,1000],z1,Spindle \WObj:=Deburring;
		MoveL [[25.282,28.339,56.857],[0.18935116,0.68232004,-0.68128306,0.18557723],[-1,0,-1,0],[9E+09,9E+09,9E+09,9E+09,9E+09,9E+09]],[16.67,500,5000,1000],z1,Spindle \WObj:=Deburring;
		MoveL [[25.684,28.319,56.871],[0.18522154,0.68111918,-0.68241816,0.18993444],[-1,0,-1,0],[9E+09,9E+09,9E+09,9E+09,9E+09,9E+09]],[16.67,500,5000,1000],z1,Spindle \WObj:=Deburring;
		MoveL [[26.080,28.259,56.914],[0.18073243,0.67999960,-0.68361950,0.19390901],[-1,-1,-1,0],[9E+09,9E+09,9E+09,9E+09,9E+09,9E+09]],[16.67,500,5000,1000],z1,Spindle \WObj:=Deburring;
		MoveL [[26.465,28.160,56.985],[0.17623862,0.67888710,-0.68479209,0.19776767],[-1,-1,-1,0],[9E+09,9E+09,9E+09,9E+09,9E+09,9E+09]],[16.67,500,5000,1000],z1,Spindle \WObj:=Deburring;
		MoveL [[26.831,28.024,57.082],[0.17210736,0.67764653,-0.68584188,0.20197810],[-1,-1,-1,0],[9E+09,9E+09,9E+09,9E+09,9E+09,9E+09]],[16.67,500,5000,1000],z1,Spindle \WObj:=Deburring;
		MoveL [[27.175,27.852,57.206],[0.16912286,0.67631769,-0.68658532,0.20637936],[-1,-1,-1,0],[9E+09,9E+09,9E+09,9E+09,9E+09,9E+09]],[16.67,500,5000,1000],z1,Spindle \WObj:=Deburring;
		MoveL [[27.490,27.648,57.352],[0.16776395,0.67481575,-0.68691632,0.21124613],[-1,-1,-1,0],[9E+09,9E+09,9E+09,9E+09,9E+09,9E+09]],[16.67,500,5000,1000],z1,Spindle \WObj:=Deburring;
		MoveL [[27.771,27.413,57.521],[0.16798658,0.67321581,-0.68686149,0.21629208],[-1,-1,-1,0],[9E+09,9E+09,9E+09,9E+09,9E+09,9E+09]],[16.67,500,5000,1000],z1,Spindle \WObj:=Deburring;
		MoveL [[28.016,27.152,57.708],[0.16815382,0.67155917,-0.68682051,0.22138237],[0,-1,-1,0],[9E+09,9E+09,9E+09,9E+09,9E+09,9E+09]],[16.67,500,5000,1000],z1,Spindle \WObj:=Deburring;
		MoveL [[28.222,26.870,57.909],[0.16787842,0.66975932,-0.68688902,0.22676588],[0,-1,-1,0],[9E+09,9E+09,9E+09,9E+09,9E+09,9E+09]],[16.67,500,5000,1000],z1,Spindle \WObj:=Deburring;
		MoveL [[28.384,26.569,58.122],[0.16741010,0.66790825,-0.68700485,0.23215674],[0,-1,-1,0],[9E+09,9E+09,9E+09,9E+09,9E+09,9E+09]],[16.67,500,5000,1000],z1,Spindle \WObj:=Deburring;
		MoveL [[28.501,26.253,58.345],[0.16734901,0.66607097,-0.68701935,0.23737771],[0,-1,-1,0],[9E+09,9E+09,9E+09,9E+09,9E+09,9E+09]],[16.67,500,5000,1000],z1,Spindle \WObj:=Deburring;
		MoveL [[28.572,25.928,58.573],[0.16786760,0.66426426,-0.68689039,0.24239443],[0,-1,0,0],[9E+09,9E+09,9E+09,9E+09,9E+09,9E+09]],[16.67,500,5000,1000],z1,Spindle \WObj:=Deburring;
		MoveL [[28.596,25.599,58.803],[0.16910296,0.66265114,-0.68658797,0.24676836],[0,-1,0,0],[9E+09,9E+09,9E+09,9E+09,9E+09,9E+09]],[16.67,500,5000,1000],z1,Spindle \WObj:=Deburring;
		MoveL [[28.572,25.269,59.034],[0.17202286,0.66150771,-0.68586326,0.24981447],[0,-1,0,0],[9E+09,9E+09,9E+09,9E+09,9E+09,9E+09]],[16.67,500,5000,1000],z1,Spindle \WObj:=Deburring;
		MoveL [[28.501,24.943,59.260],[0.17639119,0.66090829,-0.68475329,0.25139474],[0,-1,-1,0],[9E+09,9E+09,9E+09,9E+09,9E+09,9E+09]],[16.67,500,5000,1000],z1,Spindle \WObj:=Deburring;
		MoveL [[28.384,24.625,59.480],[0.18152823,0.66067877,-0.68340711,0.25200355],[0,-1,-1,0],[9E+09,9E+09,9E+09,9E+09,9E+09,9E+09]],[16.67,500,5000,1000],z1,Spindle \WObj:=Deburring;
		MoveL [[28.222,24.321,59.689],[0.18692983,0.66037836,-0.68195084,0.25278590],[0,-1,-1,0],[9E+09,9E+09,9E+09,9E+09,9E+09,9E+09]],[16.67,500,5000,1000],z1,Spindle \WObj:=Deburring;
		MoveL [[28.018,24.033,59.884],[0.19150685,0.65987166,-0.68067884,0.25410791],[0,-1,-1,0],[9E+09,9E+09,9E+09,9E+09,9E+09,9E+09]],[16.67,500,5000,1000],z1,Spindle \WObj:=Deburring;
		MoveL [[27.774,23.767,60.064],[0.19658865,0.65953389,-0.67923044,0.25497836],[0,-1,-1,0],[9E+09,9E+09,9E+09,9E+09,9E+09,9E+09]],[16.67,500,5000,1000],z1,Spindle \WObj:=Deburring;
		MoveL [[27.492,23.528,60.225],[0.20152635,0.65948841,-0.67778057,0.25509932],[0,-1,-1,0],[9E+09,9E+09,9E+09,9E+09,9E+09,9E+09]],[16.67,500,5000,1000],z1,Spindle \WObj:=Deburring;
		MoveL [[27.178,23.317,60.366],[0.20658164,0.65986226,-0.67625713,0.25413014],[0,-1,-1,0],[9E+09,9E+09,9E+09,9E+09,9E+09,9E+09]],[16.67,500,5000,1000],z1,Spindle \WObj:=Deburring;
		MoveL [[26.836,23.140,60.484],[0.21165497,0.66080736,-0.67468503,0.25166629],[-1,-1,-1,0],[9E+09,9E+09,9E+09,9E+09,9E+09,9E+09]],[16.67,500,5000,1000],z1,Spindle \WObj:=Deburring;
		MoveL [[26.470,22.999,60.579],[0.21641718,0.66238591,-0.67317454,0.24747636],[-1,-1,-1,0],[9E+09,9E+09,9E+09,9E+09,9E+09,9E+09]],[16.67,500,5000,1000],z1,Spindle \WObj:=Deburring;
		MoveL [[26.185,22.915,60.635],[0.21841829,0.66354541,-0.67252922,0.24434686],[-1,-1,-1,0],[9E+09,9E+09,9E+09,9E+09,9E+09,9E+09]],[16.67,500,5000,1000],z1,Spindle \WObj:=Deburring;
		MoveL [[25.791,22.842,60.684],[0.22302303,0.66531110,-0.67101637,0.23949720],[-1,-1,-1,0],[9E+09,9E+09,9E+09,9E+09,9E+09,9E+09]],[16.67,500,5000,1000],z1,Spindle \WObj:=Deburring;
		MoveL [[25.702,22.835,60.689],[0.22584907,0.66602478,-0.67007066,0.23750474],[-1,-1,-1,0],[9E+09,9E+09,9E+09,9E+09,9E+09,9E+09]],[16.67,500,5000,1000],z1,Spindle \WObj:=Deburring;
		MoveL [[25.612,22.828,60.693],[0.22589446,0.66594179,-0.67005520,0.23773778],[-1,-1,-1,0],[9E+09,9E+09,9E+09,9E+09,9E+09,9E+09]],[16.67,500,5000,1000],z1,Spindle \WObj:=Deburring;
		MoveL [[25.523,22.821,60.698],[0.22593931,0.66585901,-0.67003984,0.23797020],[-1,-1,-1,0],[9E+09,9E+09,9E+09,9E+09,9E+09,9E+09]],[16.67,500,5000,1000],z1,Spindle \WObj:=Deburring;
		MoveL [[25.494,22.829,60.691],[0.22593931,0.66585901,-0.67003984,0.23797020],[-1,-1,-1,0],[9E+09,9E+09,9E+09,9E+09,9E+09,9E+09]],[16.67,500,5000,1000],z1,Spindle \WObj:=Deburring;
		MoveL [[25.481,22.851,60.674],[0.22593931,0.66585901,-0.67003984,0.23797020],[-1,-1,-1,0],[9E+09,9E+09,9E+09,9E+09,9E+09,9E+09]],[16.67,500,5000,1000],z1,Spindle \WObj:=Deburring;
		MoveL [[25.461,22.869,60.659],[0.22593931,0.66585901,-0.67003984,0.23797020],[-1,-1,-1,0],[9E+09,9E+09,9E+09,9E+09,9E+09,9E+09]],[16.67,500,5000,1000],z1,Spindle \WObj:=Deburring;
		MoveL [[25.443,22.893,60.655],[0.22593931,0.66585901,-0.67003984,0.23797020],[-1,-1,-1,0],[9E+09,9E+09,9E+09,9E+09,9E+09,9E+09]],[16.67,500,5000,1000],z1,Spindle \WObj:=Deburring;
		MoveL [[25.435,22.918,60.671],[0.22593931,0.66585901,-0.67003984,0.23797020],[-1,-1,-1,0],[9E+09,9E+09,9E+09,9E+09,9E+09,9E+09]],[16.67,500,5000,1000],z1,Spindle \WObj:=Deburring;
		MoveL [[25.420,23.566,61.492],[0.22593931,0.66585901,-0.67003984,0.23797020],[-1,-1,-1,0],[9E+09,9E+09,9E+09,9E+09,9E+09,9E+09]],v1000,z1,Spindle \WObj:=Deburring;
		MoveL [[25.420,23.566,86.000],[0.22593931,0.66585901,-0.67003984,0.23797020],[-1,-1,-1,0],[9E+09,9E+09,9E+09,9E+09,9E+09,9E+09]],v1000,z1,Spindle \WObj:=Deburring;
		TPWrite "/'NEW SECTION'";
		TPWrite "/'Strategy: swarf5d'";
		TPWrite "/'Comment: Swarf10'";
		TPWrite "/'MATRIX DEFINITION'";
		TPWrite "/'Output x(i),y(i),z(i)'";
		TPWrite "/'Output x(j),y(j),z(j)'";
		TPWrite "/'Output x(k),y(k),z(k)'";
		TPWrite "/'Output dx,dy,dz'";
		SetTool 3;
		SetRPM 5000.0;
		MoveL [[25.692,45.602,86.000],[0.13216059,0.69456868,-0.69464675,0.13256630],[-1,0,-1,0],[9E+09,9E+09,9E+09,9E+09,9E+09,9E+09]],v1000,z1,Spindle \WObj:=Deburring;
		MoveL [[25.692,45.602,46.600],[0.13216059,0.69456868,-0.69464675,0.13256630],[-1,0,-1,0],[9E+09,9E+09,9E+09,9E+09,9E+09,9E+09]],v1000,z1,Spindle \WObj:=Deburring;
		MoveL [[25.693,45.209,45.608],[0.13216059,0.69456868,-0.69464675,0.13256630],[-1,0,-1,0],[9E+09,9E+09,9E+09,9E+09,9E+09,9E+09]],[16.67,500,5000,1000],z1,Spindle \WObj:=Deburring;
		MoveL [[25.702,45.206,45.579],[0.13216059,0.69456868,-0.69464675,0.13256630],[-1,0,-1,0],[9E+09,9E+09,9E+09,9E+09,9E+09,9E+09]],[16.67,500,5000,1000],z1,Spindle \WObj:=Deburring;
		MoveL [[25.723,45.219,45.561],[0.13216059,0.69456868,-0.69464675,0.13256630],[-1,0,-1,0],[9E+09,9E+09,9E+09,9E+09,9E+09,9E+09]],[16.67,500,5000,1000],z1,Spindle \WObj:=Deburring;
		MoveL [[25.747,45.239,45.554],[0.13216059,0.69456868,-0.69464675,0.13256630],[-1,0,-1,0],[9E+09,9E+09,9E+09,9E+09,9E+09,9E+09]],[16.67,500,5000,1000],z1,Spindle \WObj:=Deburring;
		MoveL [[25.764,45.263,45.545],[0.13216059,0.69456868,-0.69464675,0.13256630],[-1,0,-1,0],[9E+09,9E+09,9E+09,9E+09,9E+09,9E+09]],[16.67,500,5000,1000],z1,Spindle \WObj:=Deburring;
		MoveL [[25.794,45.268,45.543],[0.13216059,0.69456868,-0.69464675,0.13256630],[-1,0,-1,0],[9E+09,9E+09,9E+09,9E+09,9E+09,9E+09]],[16.67,500,5000,1000],z1,Spindle \WObj:=Deburring;
		MoveL [[26.025,45.228,45.565],[0.12884607,0.69348474,-0.69526762,0.13813234],[-1,0,-1,0],[9E+09,9E+09,9E+09,9E+09,9E+09,9E+09]],[16.67,500,5000,1000],z1,Spindle \WObj:=Deburring;
		MoveL [[26.411,45.122,45.621],[0.12743080,0.69192899,-0.69552998,0.14571789],[-1,-1,-1,0],[9E+09,9E+09,9E+09,9E+09,9E+09,9E+09]],[16.67,500,5000,1000],z1,Spindle \WObj:=Deburring;
		MoveL [[26.690,45.018,45.676],[0.12817009,0.69085540,-0.69539292,0.15073133],[-1,-1,-1,0],[9E+09,9E+09,9E+09,9E+09,9E+09,9E+09]],[16.67,500,5000,1000],z1,Spindle \WObj:=Deburring;
		MoveL [[27.042,44.841,45.770],[0.12762693,0.68907449,-0.69549355,0.15867080],[-1,-1,-1,0],[9E+09,9E+09,9E+09,9E+09,9E+09,9E+09]],[16.67,500,5000,1000],z1,Spindle \WObj:=Deburring;
		MoveL [[27.366,44.628,45.884],[0.12659289,0.68725464,-0.69568116,0.16638217],[-1,-1,-1,0],[9E+09,9E+09,9E+09,9E+09,9E+09,9E+09]],[16.67,500,5000,1000],z1,Spindle \WObj:=Deburring;
		MoveL [[27.685,44.359,46.029],[0.12656719,0.68523255,-0.69568718,0.17451777],[-1,-1,-1,0],[9E+09,9E+09,9E+09,9E+09,9E+09,9E+09]],[16.67,500,5000,1000],z1,Spindle \WObj:=Deburring;
		MoveL [[27.992,44.007,46.221],[0.12813389,0.68264677,-0.69540084,0.18437126],[0,-1,-1,0],[9E+09,9E+09,9E+09,9E+09,9E+09,9E+09]],[16.67,500,5000,1000],z1,Spindle \WObj:=Deburring;
		MoveL [[28.198,43.704,46.391],[0.12981649,0.68090681,-0.69508732,0.19070186],[0,-1,0,0],[9E+09,9E+09,9E+09,9E+09,9E+09,9E+09]],[16.67,500,5000,1000],z1,Spindle \WObj:=Deburring;
		MoveL [[28.364,43.383,46.572],[0.13277788,0.67923932,-0.69452861,0.19655534],[0,-1,0,0],[9E+09,9E+09,9E+09,9E+09,9E+09,9E+09]],[16.67,500,5000,1000],z1,Spindle \WObj:=Deburring;
		MoveL [[28.485,43.049,46.765],[0.13669254,0.67766392,-0.69376890,0.20191948],[0,-1,0,0],[9E+09,9E+09,9E+09,9E+09,9E+09,9E+09]],[16.67,500,5000,1000],z1,Spindle \WObj:=Deburring;
		MoveL [[28.564,42.706,46.965],[0.14094340,0.67605961,-0.69291804,0.20722682],[0,-1,0,0],[9E+09,9E+09,9E+09,9E+09,9E+09,9E+09]],[16.67,500,5000,1000],z1,Spindle \WObj:=Deburring;
		MoveL [[28.596,42.360,47.170],[0.14491289,0.67422403,-0.69209870,0.21312343],[0,-1,0,0],[9E+09,9E+09,9E+09,9E+09,9E+09,9E+09]],[16.67,500,5000,1000],z1,Spindle \WObj:=Deburring;
		MoveL [[28.581,42.013,47.377],[0.14828967,0.67220222,-0.69138353,0.21941551],[0,-1,0,0],[9E+09,9E+09,9E+09,9E+09,9E+09,9E+09]],[16.67,500,5000,1000],z1,Spindle \WObj:=Deburring;
		MoveL [[28.521,41.671,47.584],[0.15110433,0.66986910,-0.69077246,0.22644267],[0,-1,0,0],[9E+09,9E+09,9E+09,9E+09,9E+09,9E+09]],[16.67,500,5000,1000],z1,Spindle \WObj:=Deburring;
		MoveL [[28.414,41.339,47.787],[0.15466273,0.66765208,-0.68998605,0.23289355],[0,-1,0,0],[9E+09,9E+09,9E+09,9E+09,9E+09,9E+09]],[16.67,500,5000,1000],z1,Spindle \WObj:=Deburring;
		MoveL [[28.264,41.020,47.985],[0.15922818,0.66573189,-0.68894409,0.23833479],[0,-1,0,0],[9E+09,9E+09,9E+09,9E+09,9E+09,9E+09]],[16.67,500,5000,1000],z1,Spindle \WObj:=Deburring;
		MoveL [[28.070,40.719,48.173],[0.16493912,0.66412244,-0.68759962,0.24278229],[0,-1,0,0],[9E+09,9E+09,9E+09,9E+09,9E+09,9E+09]],[16.67,500,5000,1000],z1,Spindle \WObj:=Deburring;
		MoveL [[27.902,40.506,48.308],[0.16843127,0.66316504,-0.68675428,0.24538050],[0,-1,0,0],[9E+09,9E+09,9E+09,9E+09,9E+09,9E+09]],[16.67,500,5000,1000],z1,Spindle \WObj:=Deburring;
		MoveL [[27.613,40.225,48.488],[0.17621526,0.66230241,-0.68479880,0.24769800],[0,-1,-1,0],[9E+09,9E+09,9E+09,9E+09,9E+09,9E+09]],[16.67,500,5000,1000],z1,Spindle \WObj:=Deburring;
		MoveL [[27.311,39.999,48.633],[0.18399084,0.66224732,-0.68274923,0.24784945],[0,-1,-1,0],[9E+09,9E+09,9E+09,9E+09,9E+09,9E+09]],[16.67,500,5000,1000],z1,Spindle \WObj:=Deburring;
		MoveL [[26.979,39.805,48.759],[0.19203488,0.66164443,-0.68053091,0.24945328],[0,-1,-1,0],[9E+09,9E+09,9E+09,9E+09,9E+09,9E+09]],[16.67,500,5000,1000],z1,Spindle \WObj:=Deburring;
		MoveL [[26.621,39.646,48.861],[0.20041228,0.66114167,-0.67811139,0.25078189],[0,-1,-1,0],[9E+09,9E+09,9E+09,9E+09,9E+09,9E+09]],[16.67,500,5000,1000],z1,Spindle \WObj:=Deburring;
		MoveL [[26.242,39.526,48.938],[0.20887227,0.66118185,-0.67555415,0.25067415],[-1,-1,-1,0],[9E+09,9E+09,9E+09,9E+09,9E+09,9E+09]],[16.67,500,5000,1000],z1,Spindle \WObj:=Deburring;
		MoveL [[25.849,39.446,48.990],[0.21701095,0.66191240,-0.67298126,0.24874573],[-1,-1,-1,0],[9E+09,9E+09,9E+09,9E+09,9E+09,9E+09]],[16.67,500,5000,1000],z1,Spindle \WObj:=Deburring;
		MoveL [[25.447,39.407,49.016],[0.22466021,0.66330398,-0.67046930,0.24500315],[-1,-1,-1,0],[9E+09,9E+09,9E+09,9E+09,9E+09,9E+09]],[16.67,500,5000,1000],z1,Spindle \WObj:=Deburring;
		MoveL [[24.943,39.424,49.005],[0.23279172,0.66652871,-0.66768994,0.23608818],[-1,0,-1,0],[9E+09,9E+09,9E+09,9E+09,9E+09,9E+09]],[16.67,500,5000,1000],z1,Spindle \WObj:=Deburring;
		MoveL [[24.544,39.481,48.969],[0.23714323,0.66907009,-0.66615722,0.22878562],[-1,0,-1,0],[9E+09,9E+09,9E+09,9E+09,9E+09,9E+09]],[16.67,500,5000,1000],z1,Spindle \WObj:=Deburring;
		MoveL [[24.158,39.579,48.905],[0.24017855,0.67177607,-0.66506895,0.22071355],[-1,0,-1,0],[9E+09,9E+09,9E+09,9E+09,9E+09,9E+09]],[16.67,500,5000,1000],z1,Spindle \WObj:=Deburring;
		MoveL [[23.788,39.717,48.816],[0.24263839,0.67438671,-0.66417192,0.21261428],[-1,0,-1,0],[9E+09,9E+09,9E+09,9E+09,9E+09,9E+09]],[16.67,500,5000,1000],z1,Spindle \WObj:=Deburring;
		MoveL [[23.441,39.890,48.704],[0.24476623,0.67682827,-0.66339072,0.20470891],[-1,0,-1,0],[9E+09,9E+09,9E+09,9E+09,9E+09,9E+09]],[16.67,500,5000,1000],z1,Spindle \WObj:=Deburring;
		MoveL [[23.197,40.041,48.607],[0.24540922,0.67816539,-0.66315559,0.20022657],[-1,0,-1,0],[9E+09,9E+09,9E+09,9E+09,9E+09,9E+09]],[16.67,500,5000,1000],z1,Spindle \WObj:=Deburring;
		MoveL [[22.876,40.296,48.443],[0.24464096,0.68061402,-0.66343796,0.19174312],[-1,0,-1,0],[9E+09,9E+09,9E+09,9E+09,9E+09,9E+09]],[16.67,500,5000,1000],z1,Spindle \WObj:=Deburring;
		MoveL [[22.567,40.633,48.229],[0.24315224,0.68352168,-0.66398726,0.18109671],[-1,0,-1,0],[9E+09,9E+09,9E+09,9E+09,9E+09,9E+09]],[16.67,500,5000,1000],z1,Spindle \WObj:=Deburring;
		MoveL [[22.360,40.927,48.043],[0.24201463,0.68532578,-0.66439950,0.17415737],[-1,0,-1,0],[9E+09,9E+09,9E+09,9E+09,9E+09,9E+09]],[16.67,500,5000,1000],z1,Spindle \WObj:=Deburring;
		MoveL [[22.197,41.240,47.848],[0.23982955,0.68690232,-0.66519351,0.16782307],[-1,0,-1,0],[9E+09,9E+09,9E+09,9E+09,9E+09,9E+09]],[16.67,500,5000,1000],z1,Spindle \WObj:=Deburring;
		MoveL [[22.077,41.569,47.645],[0.23642676,0.68821274,-0.66640941,0.16237028],[-1,0,-1,0],[9E+09,9E+09,9E+09,9E+09,9E+09,9E+09]],[16.67,500,5000,1000],z1,Spindle \WObj:=Deburring;
		MoveL [[22.002,41.908,47.439],[0.23198967,0.68933999,-0.66796683,0.15751661],[-1,0,-1,0],[9E+09,9E+09,9E+09,9E+09,9E+09,9E+09]],[16.67,500,5000,1000],z1,Spindle \WObj:=Deburring;
		MoveL [[21.973,42.254,47.232],[0.22705063,0.69031417,-0.66966357,0.15318312],[-1,0,-1,0],[9E+09,9E+09,9E+09,9E+09,9E+09,9E+09]],[16.67,500,5000,1000],z1,Spindle \WObj:=Deburring;
		MoveL [[21.992,42.601,47.026],[0.22127466,0.69107431,-0.67159198,0.14972652],[-1,0,-1,0],[9E+09,9E+09,9E+09,9E+09,9E+09,9E+09]],[16.67,500,5000,1000],z1,Spindle \WObj:=Deburring;
		MoveL [[22.056,42.946,46.825],[0.21568812,0.69193435,-0.67340807,0.14569513],[-1,0,-1,0],[9E+09,9E+09,9E+09,9E+09,9E+09,9E+09]],[16.67,500,5000,1000],z1,Spindle \WObj:=Deburring;
		MoveL [[22.165,43.283,46.631],[0.21018080,0.69285953,-0.67514594,0.14123620],[-1,0,-1,0],[9E+09,9E+09,9E+09,9E+09,9E+09,9E+09]],[16.67,500,5000,1000],z1,Spindle \WObj:=Deburring;
		MoveL [[22.317,43.608,46.445],[0.20471438,0.69386364,-0.67682510,0.13620959],[-1,0,-1,0],[9E+09,9E+09,9E+09,9E+09,9E+09,9E+09]],[16.67,500,5000,1000],z1,Spindle \WObj:=Deburring;
		MoveL [[22.510,43.918,46.271],[0.19897401,0.69490073,-0.67853492,0.13081545],[-1,0,-1,0],[9E+09,9E+09,9E+09,9E+09,9E+09,9E+09]],[16.67,500,5000,1000],z1,Spindle \WObj:=Deburring;
		MoveL [[22.678,44.139,46.148],[0.19557188,0.69558560,-0.67952234,0.12712868],[-1,0,-1,0],[9E+09,9E+09,9E+09,9E+09,9E+09,9E+09]],[16.67,500,5000,1000],z1,Spindle \WObj:=Deburring;
		MoveL [[22.965,44.433,45.988],[0.18811326,0.69625403,-0.68162473,0.12341581],[-1,0,-1,0],[9E+09,9E+09,9E+09,9E+09,9E+09,9E+09]],[16.67,500,5000,1000],z1,Spindle \WObj:=Deburring;
		MoveL [[23.265,44.672,45.859],[0.18090936,0.69646069,-0.68357353,0.12223564],[-1,0,-1,0],[9E+09,9E+09,9E+09,9E+09,9E+09,9E+09]],[16.67,500,5000,1000],z1,Spindle \WObj:=Deburring;
		MoveL [[23.595,44.878,45.749],[0.17344619,0.69663471,-0.68550400,0.12124674],[-1,0,-1,0],[9E+09,9E+09,9E+09,9E+09,9E+09,9E+09]],[16.67,500,5000,1000],z1,Spindle \WObj:=Deburring;
		MoveL [[23.951,45.048,45.660],[0.16576860,0.69660157,-0.68740202,0.12143102],[-1,0,-1,0],[9E+09,9E+09,9E+09,9E+09,9E+09,9E+09]],[16.67,500,5000,1000],z1,Spindle \WObj:=Deburring;
		MoveL [[24.328,45.178,45.592],[0.15776477,0.69643808,-0.68928166,0.12237267],[-1,0,-1,0],[9E+09,9E+09,9E+09,9E+09,9E+09,9E+09]],[16.67,500,5000,1000],z1,Spindle \WObj:=Deburring;
		MoveL [[24.721,45.266,45.546],[0.14927369,0.69628878,-0.69117005,0.12322040],[-1,0,-1,0],[9E+09,9E+09,9E+09,9E+09,9E+09,9E+09]],[16.67,500,5000,1000],z1,Spindle \WObj:=Deburring;
		MoveL [[25.122,45.307,45.523],[0.14133769,0.69587357,-0.69283837,0.12553337],[-1,0,-1,0],[9E+09,9E+09,9E+09,9E+09,9E+09,9E+09]],[16.67,500,5000,1000],z1,Spindle \WObj:=Deburring;
		MoveL [[25.616,45.291,45.532],[0.13276073,0.69468731,-0.69453115,0.13194930],[-1,0,-1,0],[9E+09,9E+09,9E+09,9E+09,9E+09,9E+09]],[16.67,500,5000,1000],z1,Spindle \WObj:=Deburring;
		MoveL [[25.705,45.279,45.538],[0.13246067,0.69462776,-0.69458933,0.13225770],[-1,0,-1,0],[9E+09,9E+09,9E+09,9E+09,9E+09,9E+09]],[16.67,500,5000,1000],z1,Spindle \WObj:=Deburring;
		MoveL [[25.794,45.268,45.543],[0.13216059,0.69456868,-0.69464675,0.13256630],[-1,0,-1,0],[9E+09,9E+09,9E+09,9E+09,9E+09,9E+09]],[16.67,500,5000,1000],z1,Spindle \WObj:=Deburring;
		MoveL [[25.820,45.253,45.550],[0.13216059,0.69456868,-0.69464675,0.13256630],[-1,0,-1,0],[9E+09,9E+09,9E+09,9E+09,9E+09,9E+09]],[16.67,500,5000,1000],z1,Spindle \WObj:=Deburring;
		MoveL [[25.826,45.225,45.561],[0.13216059,0.69456868,-0.69464675,0.13256630],[-1,0,-1,0],[9E+09,9E+09,9E+09,9E+09,9E+09,9E+09]],[16.67,500,5000,1000],z1,Spindle \WObj:=Deburring;
		MoveL [[25.840,45.199,45.572],[0.13216059,0.69456868,-0.69464675,0.13256630],[-1,0,-1,0],[9E+09,9E+09,9E+09,9E+09,9E+09,9E+09]],[16.67,500,5000,1000],z1,Spindle \WObj:=Deburring;
		MoveL [[25.839,45.609,46.608],[0.13216059,0.69456868,-0.69464675,0.13256630],[-1,0,-1,0],[9E+09,9E+09,9E+09,9E+09,9E+09,9E+09]],v1000,z1,Spindle \WObj:=Deburring;
		MoveL [[25.839,45.609,86.000],[0.13216059,0.69456868,-0.69464675,0.13256630],[-1,0,-1,0],[9E+09,9E+09,9E+09,9E+09,9E+09,9E+09]],v1000,z1,Spindle \WObj:=Deburring;
		TPWrite "/'NEW SECTION'";
		TPWrite "/'Strategy: swarf5d'";
		TPWrite "/'Comment: Swarf11'";
		TPWrite "/'MATRIX DEFINITION'";
		TPWrite "/'Output x(i),y(i),z(i)'";
		TPWrite "/'Output x(j),y(j),z(j)'";
		TPWrite "/'Output x(k),y(k),z(k)'";
		TPWrite "/'Output dx,dy,dz'";
		SetTool 3;
		SetRPM 5000.0;
		MoveL [[-52.281,-78.443,86.000],[0.04865817,0.69827538,-0.70543105,0.11140424],[0,-1,0,0],[9E+09,9E+09,9E+09,9E+09,9E+09,9E+09]],v1000,z1,Spindle \WObj:=Deburring;
		MoveL [[-52.281,-78.443,22.215],[0.04865817,0.69827538,-0.70543105,0.11140424],[0,-1,0,0],[9E+09,9E+09,9E+09,9E+09,9E+09,9E+09]],v1000,z1,Spindle \WObj:=Deburring;
		MoveL [[-52.063,-79.007,19.782],[0.04865817,0.69827538,-0.70543105,0.11140424],[0,-1,0,0],[9E+09,9E+09,9E+09,9E+09,9E+09,9E+09]],[16.67,500,5000,1000],z1,Spindle \WObj:=Deburring;
		MoveL [[-51.845,-79.572,17.349],[0.04865817,0.69827538,-0.70543105,0.11140424],[0,-1,0,0],[9E+09,9E+09,9E+09,9E+09,9E+09,9E+09]],[16.67,500,5000,1000],z1,Spindle \WObj:=Deburring;
		MoveL [[-51.831,-79.570,17.319],[0.04865817,0.69827538,-0.70543105,0.11140424],[0,-1,0,0],[9E+09,9E+09,9E+09,9E+09,9E+09,9E+09]],[16.67,500,5000,1000],z1,Spindle \WObj:=Deburring;
		MoveL [[-51.805,-79.554,17.307],[0.04865817,0.69827538,-0.70543105,0.11140424],[0,-1,0,0],[9E+09,9E+09,9E+09,9E+09,9E+09,9E+09]],[16.67,500,5000,1000],z1,Spindle \WObj:=Deburring;
		MoveL [[-51.780,-79.534,17.309],[0.04865817,0.69827538,-0.70543105,0.11140424],[0,-1,0,0],[9E+09,9E+09,9E+09,9E+09,9E+09,9E+09]],[16.67,500,5000,1000],z1,Spindle \WObj:=Deburring;
		MoveL [[-51.752,-79.523,17.312],[0.04865817,0.69827538,-0.70543105,0.11140424],[0,-1,0,0],[9E+09,9E+09,9E+09,9E+09,9E+09,9E+09]],[16.67,500,5000,1000],z1,Spindle \WObj:=Deburring;
		MoveL [[-51.740,-79.494,17.313],[0.04865817,0.69827538,-0.70543105,0.11140424],[0,-1,0,0],[9E+09,9E+09,9E+09,9E+09,9E+09,9E+09]],[16.67,500,5000,1000],z1,Spindle \WObj:=Deburring;
		MoveL [[-51.740,-74.500,17.313],[0.04638831,0.69863571,-0.70558269,0.10912989],[0,-1,0,0],[9E+09,9E+09,9E+09,9E+09,9E+09,9E+09]],[16.67,500,5000,1000],z1,Spindle \WObj:=Deburring;
		MoveL [[-51.740,-69.507,17.313],[0.04412570,0.69898771,-0.70572861,0.10684671],[0,-1,0,0],[9E+09,9E+09,9E+09,9E+09,9E+09,9E+09]],[16.67,500,5000,1000],z1,Spindle \WObj:=Deburring;
		MoveL [[-51.739,-64.513,17.313],[0.04185805,0.69933280,-0.70586632,0.10456710],[0,-1,0,0],[9E+09,9E+09,9E+09,9E+09,9E+09,9E+09]],[16.67,500,5000,1000],z1,Spindle \WObj:=Deburring;
		MoveL [[-51.739,-59.519,17.313],[0.03959158,0.69966993,-0.70599738,0.10228489],[0,-1,0,0],[9E+09,9E+09,9E+09,9E+09,9E+09,9E+09]],[16.67,500,5000,1000],z1,Spindle \WObj:=Deburring;
		MoveL [[-51.739,-54.525,17.313],[0.03732611,0.70000033,-0.70612057,0.10000018],[0,-1,0,0],[9E+09,9E+09,9E+09,9E+09,9E+09,9E+09]],[16.67,500,5000,1000],z1,Spindle \WObj:=Deburring;
		MoveL [[-51.738,-49.531,17.313],[0.03506185,0.70032277,-0.70623712,0.09771294],[0,-1,0,0],[9E+09,9E+09,9E+09,9E+09,9E+09,9E+09]],[16.67,500,5000,1000],z1,Spindle \WObj:=Deburring;
		MoveL [[-51.738,-44.537,17.313],[0.03279268,0.70063751,-0.70634620,0.09542937],[0,-1,0,0],[9E+09,9E+09,9E+09,9E+09,9E+09,9E+09]],[16.67,500,5000,1000],z1,Spindle \WObj:=Deburring;
		MoveL [[-51.738,-39.543,17.313],[0.03052396,0.70094548,-0.70644755,0.09314279],[0,-1,0,0],[9E+09,9E+09,9E+09,9E+09,9E+09,9E+09]],[16.67,500,5000,1000],z1,Spindle \WObj:=Deburring;
		MoveL [[-51.737,-34.549,17.313],[0.02825715,0.70124539,-0.70654222,0.09085445],[0,-1,0,0],[9E+09,9E+09,9E+09,9E+09,9E+09,9E+09]],[16.67,500,5000,1000],z1,Spindle \WObj:=Deburring;
		MoveL [[-51.737,-29.555,17.313],[0.02599113,0.70153850,-0.70662911,0.08856347],[0,-1,0,0],[9E+09,9E+09,9E+09,9E+09,9E+09,9E+09]],[16.67,500,5000,1000],z1,Spindle \WObj:=Deburring;
		MoveL [[-51.737,-24.561,17.313],[0.02372020,0.70182377,-0.70670868,0.08627623],[0,-1,0,0],[9E+09,9E+09,9E+09,9E+09,9E+09,9E+09]],[16.67,500,5000,1000],z1,Spindle \WObj:=Deburring;
		MoveL [[-51.736,-19.567,17.313],[0.02145047,0.70210155,-0.70678110,0.08398669],[0,-1,0,0],[9E+09,9E+09,9E+09,9E+09,9E+09,9E+09]],[16.67,500,5000,1000],z1,Spindle \WObj:=Deburring;
		MoveL [[-51.736,-14.573,17.313],[0.01918191,0.70237185,-0.70684637,0.08169482],[0,-1,0,0],[9E+09,9E+09,9E+09,9E+09,9E+09,9E+09]],[16.67,500,5000,1000],z1,Spindle \WObj:=Deburring;
		MoveL [[-51.736,-9.579,17.313],[0.01691459,0.70263403,-0.70690512,0.07940064],[0,-1,0,0],[9E+09,9E+09,9E+09,9E+09,9E+09,9E+09]],[16.67,500,5000,1000],z1,Spindle \WObj:=Deburring;
		MoveL [[-51.735,-4.585,17.313],[0.01464226,0.70288945,-0.70695546,0.07711037],[0,-1,0,0],[9E+09,9E+09,9E+09,9E+09,9E+09,9E+09]],[16.67,500,5000,1000],z1,Spindle \WObj:=Deburring;
		MoveL [[-51.735,0.409,17.313],[0.01237120,0.70313731,-0.70699869,0.07481792],[0,-1,0,0],[9E+09,9E+09,9E+09,9E+09,9E+09,9E+09]],[16.67,500,5000,1000],z1,Spindle \WObj:=Deburring;
		MoveL [[-51.734,5.403,17.313],[0.01010144,0.70337762,-0.70703483,0.07252333],[0,-1,0,0],[9E+09,9E+09,9E+09,9E+09,9E+09,9E+09]],[16.67,500,5000,1000],z1,Spindle \WObj:=Deburring;
		MoveL [[-51.734,10.397,17.313],[0.00783285,0.70361097,-0.70706328,0.07022658],[0,-1,0,0],[9E+09,9E+09,9E+09,9E+09,9E+09,9E+09]],[16.67,500,5000,1000],z1,Spindle \WObj:=Deburring;
		MoveL [[-51.734,15.391,17.313],[0.00555945,0.70383618,-0.70708467,0.06793384],[0,-1,0,0],[9E+09,9E+09,9E+09,9E+09,9E+09,9E+09]],[16.67,500,5000,1000],z1,Spindle \WObj:=Deburring;
		MoveL [[-51.733,20.385,17.313],[0.00329353,0.70405373,-0.70709958,0.06563288],[0,-1,0,0],[9E+09,9E+09,9E+09,9E+09,9E+09,9E+09]],[16.67,500,5000,1000],z1,Spindle \WObj:=Deburring;
		MoveL [[-51.733,25.379,17.313],[0.00102271,0.70426432,-0.70710627,0.06333601],[0,-1,0,0],[9E+09,9E+09,9E+09,9E+09,9E+09,9E+09]],[16.67,500,5000,1000],z1,Spindle \WObj:=Deburring;
		MoveL [[-51.733,30.373,17.313],[0.00125294,-0.70446726,0.70710539,-0.06104325],[0,-1,0,0],[9E+09,9E+09,9E+09,9E+09,9E+09,9E+09]],[16.67,500,5000,1000],z1,Spindle \WObj:=Deburring;
		MoveL [[-51.732,35.367,17.313],[0.00352098,-0.70466255,0.70709802,-0.05874243],[0,-1,0,0],[9E+09,9E+09,9E+09,9E+09,9E+09,9E+09]],[16.67,500,5000,1000],z1,Spindle \WObj:=Deburring;
		MoveL [[-51.732,40.361,17.313],[0.00579389,-0.70485014,0.70708316,-0.05644572],[0,-1,0,0],[9E+09,9E+09,9E+09,9E+09,9E+09,9E+09]],[16.67,500,5000,1000],z1,Spindle \WObj:=Deburring;
		MoveL [[-51.732,45.355,17.313],[0.00805926,-0.70503072,0.70706116,-0.05414093],[0,-1,0,0],[9E+09,9E+09,9E+09,9E+09,9E+09,9E+09]],[16.67,500,5000,1000],z1,Spindle \WObj:=Deburring;
		MoveL [[-51.731,50.349,17.313],[0.01032934,-0.70520355,0.70703171,-0.05184045],[0,-1,0,0],[9E+09,9E+09,9E+09,9E+09,9E+09,9E+09]],[16.67,500,5000,1000],z1,Spindle \WObj:=Deburring;
		MoveL [[-51.731,55.343,17.313],[0.01260421,-0.70536917,0.70699423,-0.04954422],[0,-1,0,0],[9E+09,9E+09,9E+09,9E+09,9E+09,9E+09]],[16.67,500,5000,1000],z1,Spindle \WObj:=Deburring;
		MoveL [[-51.731,60.337,17.313],[0.01487143,-0.70552716,0.70695024,-0.04724000],[0,-1,0,0],[9E+09,9E+09,9E+09,9E+09,9E+09,9E+09]],[16.67,500,5000,1000],z1,Spindle \WObj:=Deburring;
		MoveL [[-51.730,65.331,17.313],[0.01714330,-0.70567729,0.70689890,-0.04494017],[0,-1,0,0],[9E+09,9E+09,9E+09,9E+09,9E+09,9E+09]],[16.67,500,5000,1000],z1,Spindle \WObj:=Deburring;
		MoveL [[-51.730,70.325,17.313],[0.01941375,-0.70582026,0.70684003,-0.04263851],[0,-1,0,0],[9E+09,9E+09,9E+09,9E+09,9E+09,9E+09]],[16.67,500,5000,1000],z1,Spindle \WObj:=Deburring;
		MoveL [[-51.730,75.319,17.313],[0.02168271,-0.70595546,0.70677425,-0.04033506],[0,-1,0,0],[9E+09,9E+09,9E+09,9E+09,9E+09,9E+09]],[16.67,500,5000,1000],z1,Spindle \WObj:=Deburring;
		MoveL [[-51.729,80.313,17.313],[0.02395009,-0.70608349,0.70670094,-0.03802996],[0,-1,0,0],[9E+09,9E+09,9E+09,9E+09,9E+09,9E+09]],[16.67,500,5000,1000],z1,Spindle \WObj:=Deburring;
		MoveL [[-51.729,85.307,17.313],[0.02622212,-0.70620352,0.70662042,-0.03572927],[0,-1,0,0],[9E+09,9E+09,9E+09,9E+09,9E+09,9E+09]],[16.67,500,5000,1000],z1,Spindle \WObj:=Deburring;
		MoveL [[-51.728,90.301,17.313],[0.02849259,-0.70631632,0.70653242,-0.03342692],[0,-1,0,0],[9E+09,9E+09,9E+09,9E+09,9E+09,9E+09]],[16.67,500,5000,1000],z1,Spindle \WObj:=Deburring;
		MoveL [[-51.728,95.295,17.313],[0.03076146,-0.70642129,0.70643758,-0.03112293],[0,-1,0,0],[9E+09,9E+09,9E+09,9E+09,9E+09,9E+09]],[16.67,500,5000,1000],z1,Spindle \WObj:=Deburring;
		MoveL [[-51.702,99.137,17.313],[0.03047199,-0.70641346,0.70645008,-0.03130140],[0,-1,0,0],[9E+09,9E+09,9E+09,9E+09,9E+09,9E+09]],[16.67,500,5000,1000],z1,Spindle \WObj:=Deburring;
		MoveL [[-51.676,102.980,17.313],[0.03018866,-0.70640524,0.70646225,-0.03148601],[0,-1,0,0],[9E+09,9E+09,9E+09,9E+09,9E+09,9E+09]],[16.67,500,5000,1000],z1,Spindle \WObj:=Deburring;
		MoveL [[-51.598,106.232,17.313],[0.02919061,-0.70636442,0.70650382,-0.03239710],[0,-1,0,0],[9E+09,9E+09,9E+09,9E+09,9E+09,9E+09]],[16.67,500,5000,1000],z1,Spindle \WObj:=Deburring;
		MoveL [[-51.513,107.752,17.313],[0.02747015,-0.70629567,0.70657311,-0.03385630],[0,-1,0,0],[9E+09,9E+09,9E+09,9E+09,9E+09,9E+09]],[16.67,500,5000,1000],z1,Spindle \WObj:=Deburring;
		MoveL [[-51.380,108.936,17.313],[0.02479565,-0.70619760,0.70667188,-0.03584654],[0,-1,0,0],[9E+09,9E+09,9E+09,9E+09,9E+09,9E+09]],[16.67,500,5000,1000],z1,Spindle \WObj:=Deburring;
		MoveL [[-51.227,109.722,17.313],[0.02140215,-0.70608753,0.70678314,-0.03794667],[0,-1,0,0],[9E+09,9E+09,9E+09,9E+09,9E+09,9E+09]],[16.67,500,5000,1000],z1,Spindle \WObj:=Deburring;
		MoveL [[-51.071,110.238,17.313],[0.01718702,-0.70597311,0.70689791,-0.04002392],[0,-1,0,0],[9E+09,9E+09,9E+09,9E+09,9E+09,9E+09]],[16.67,500,5000,1000],z1,Spindle \WObj:=Deburring;
		MoveL [[-50.911,110.638,17.313],[0.01486501,-0.70590924,0.70695033,-0.04113877],[0,-1,0,0],[9E+09,9E+09,9E+09,9E+09,9E+09,9E+09]],[16.67,500,5000,1000],z1,Spindle \WObj:=Deburring;
		MoveL [[-50.658,111.075,17.313],[0.00730773,-0.70578840,0.70706880,-0.04316292],[0,-1,0,0],[9E+09,9E+09,9E+09,9E+09,9E+09,9E+09]],[16.67,500,5000,1000],z1,Spindle \WObj:=Deburring;
		MoveL [[-50.414,111.396,17.313],[0.00166602,-0.70575515,0.70710457,-0.04370373],[0,-1,0,0],[9E+09,9E+09,9E+09,9E+09,9E+09,9E+09]],[16.67,500,5000,1000],z1,Spindle \WObj:=Deburring;
		MoveL [[-50.130,111.683,17.313],[0.00407971,0.70576574,-0.70709498,0.04352898],[0,-1,0,0],[9E+09,9E+09,9E+09,9E+09,9E+09,9E+09]],[16.67,500,5000,1000],z1,Spindle \WObj:=Deburring;
		MoveL [[-49.896,111.876,17.313],[0.00708389,0.70579719,-0.70707126,0.04301611],[0,-1,0,0],[9E+09,9E+09,9E+09,9E+09,9E+09,9E+09]],[16.67,500,5000,1000],z1,Spindle \WObj:=Deburring;
		MoveL [[-49.552,112.089,17.313],[0.01259751,0.70587067,-0.70699423,0.04179784],[0,-1,0,0],[9E+09,9E+09,9E+09,9E+09,9E+09,9E+09]],[16.67,500,5000,1000],z1,Spindle \WObj:=Deburring;
		MoveL [[-49.060,112.310,17.313],[0.01795988,0.70598359,-0.70687891,0.03983493],[0,-1,0,0],[9E+09,9E+09,9E+09,9E+09,9E+09,9E+09]],[16.67,500,5000,1000],z1,Spindle \WObj:=Deburring;
		MoveL [[-48.433,112.500,17.313],[0.02245706,0.70611003,-0.70675009,0.03753153],[0,-1,0,0],[9E+09,9E+09,9E+09,9E+09,9E+09,9E+09]],[16.67,500,5000,1000],z1,Spindle \WObj:=Deburring;
		MoveL [[-47.520,112.668,17.313],[0.02713385,0.70627647,-0.70658593,0.03425811],[0,-1,0,0],[9E+09,9E+09,9E+09,9E+09,9E+09,9E+09]],[16.67,500,5000,1000],z1,Spindle \WObj:=Deburring;
		MoveL [[-46.443,112.784,17.313],[0.02889241,0.70635505,-0.70651602,0.03260190],[0,-1,0,0],[9E+09,9E+09,9E+09,9E+09,9E+09,9E+09]],[16.67,500,5000,1000],z1,Spindle \WObj:=Deburring;
		MoveL [[-44.843,112.869,17.313],[0.03012966,0.70640797,-0.70646446,0.03143166],[0,-1,0,0],[9E+09,9E+09,9E+09,9E+09,9E+09,9E+09]],[16.67,500,5000,1000],z1,Spindle \WObj:=Deburring;
		MoveL [[-42.048,112.913,17.313],[0.03078030,0.70643407,-0.70643631,0.03084173],[0,-1,0,0],[9E+09,9E+09,9E+09,9E+09,9E+09,9E+09]],[16.67,500,5000,1000],z1,Spindle \WObj:=Deburring;
		MoveL [[-37.302,112.913,17.313],[0.03078030,0.70643407,-0.70643631,0.03084173],[0,-1,0,0],[9E+09,9E+09,9E+09,9E+09,9E+09,9E+09]],[16.67,500,5000,1000],z1,Spindle \WObj:=Deburring;
		MoveL [[-32.556,112.912,17.313],[0.03087319,0.70643740,-0.70643238,0.03076265],[0,-1,0,0],[9E+09,9E+09,9E+09,9E+09,9E+09,9E+09]],[16.67,500,5000,1000],z1,Spindle \WObj:=Deburring;
		MoveL [[-27.810,112.911,17.313],[0.03091969,0.70643906,-0.70643040,0.03072317],[0,-1,0,0],[9E+09,9E+09,9E+09,9E+09,9E+09,9E+09]],[16.67,500,5000,1000],z1,Spindle \WObj:=Deburring;
		MoveL [[-23.065,112.911,17.313],[0.03095997,0.70644099,-0.70642816,0.03068980],[0,-1,0,0],[9E+09,9E+09,9E+09,9E+09,9E+09,9E+09]],[16.67,500,5000,1000],z1,Spindle \WObj:=Deburring;
		MoveL [[-18.319,112.910,17.313],[0.03100645,0.70644202,-0.70642680,0.03065023],[0,-1,0,0],[9E+09,9E+09,9E+09,9E+09,9E+09,9E+09]],[16.67,500,5000,1000],z1,Spindle \WObj:=Deburring;
		MoveL [[-13.573,112.909,17.313],[0.03105289,0.70644368,-0.70642483,0.03061070],[0,-1,0,0],[9E+09,9E+09,9E+09,9E+09,9E+09,9E+09]],[16.67,500,5000,1000],z1,Spindle \WObj:=Deburring;
		MoveL [[-8.827,112.909,17.313],[0.03109934,0.70644532,-0.70642285,0.03057116],[0,-1,0,0],[9E+09,9E+09,9E+09,9E+09,9E+09,9E+09]],[16.67,500,5000,1000],z1,Spindle \WObj:=Deburring;
		MoveL [[-4.082,112.908,17.313],[0.03113968,0.70644724,-0.70642060,0.03053785],[0,-1,0,0],[9E+09,9E+09,9E+09,9E+09,9E+09,9E+09]],[16.67,500,5000,1000],z1,Spindle \WObj:=Deburring;
		MoveL [[0.664,112.907,17.313],[0.03118613,0.70644888,-0.70641861,0.03049831],[-1,0,-1,0],[9E+09,9E+09,9E+09,9E+09,9E+09,9E+09]],[16.67,500,5000,1000],z1,Spindle \WObj:=Deburring;
		MoveL [[5.410,112.907,17.313],[0.03123258,0.70645052,-0.70641663,0.03045877],[-1,0,-1,0],[9E+09,9E+09,9E+09,9E+09,9E+09,9E+09]],[16.67,500,5000,1000],z1,Spindle \WObj:=Deburring;
		MoveL [[10.156,112.906,17.313],[0.03127902,0.70645216,-0.70641464,0.03041924],[-1,0,-1,0],[9E+09,9E+09,9E+09,9E+09,9E+09,9E+09]],[16.67,500,5000,1000],z1,Spindle \WObj:=Deburring;
		MoveL [[14.902,112.906,17.313],[0.03131931,0.70645407,-0.70641238,0.03038587],[-1,0,-1,0],[9E+09,9E+09,9E+09,9E+09,9E+09,9E+09]],[16.67,500,5000,1000],z1,Spindle \WObj:=Deburring;
		MoveL [[19.647,112.905,17.313],[0.03136578,0.70645508,-0.70641101,0.03034630],[-1,0,-1,0],[9E+09,9E+09,9E+09,9E+09,9E+09,9E+09]],[16.67,500,5000,1000],z1,Spindle \WObj:=Deburring;
		MoveL [[24.393,112.904,17.313],[0.03141223,0.70645671,-0.70640901,0.03030677],[-1,0,-1,0],[9E+09,9E+09,9E+09,9E+09,9E+09,9E+09]],[16.67,500,5000,1000],z1,Spindle \WObj:=Deburring;
		MoveL [[29.139,112.904,17.313],[0.03145874,0.70645833,-0.70640701,0.03026729],[-1,0,-1,0],[9E+09,9E+09,9E+09,9E+09,9E+09,9E+09]],[16.67,500,5000,1000],z1,Spindle \WObj:=Deburring;
		MoveL [[33.885,112.903,17.313],[0.03149902,0.70646023,-0.70640475,0.03023392],[-1,0,-1,0],[9E+09,9E+09,9E+09,9E+09,9E+09,9E+09]],[16.67,500,5000,1000],z1,Spindle \WObj:=Deburring;
		MoveL [[38.631,112.902,17.313],[0.03154547,0.70646185,-0.70640275,0.03019439],[-1,0,-1,0],[9E+09,9E+09,9E+09,9E+09,9E+09,9E+09]],[16.67,500,5000,1000],z1,Spindle \WObj:=Deburring;
		MoveL [[43.376,112.902,17.313],[0.03159192,0.70646346,-0.70640074,0.03015486],[-1,0,-1,0],[9E+09,9E+09,9E+09,9E+09,9E+09,9E+09]],[16.67,500,5000,1000],z1,Spindle \WObj:=Deburring;
		MoveL [[45.538,112.839,17.313],[0.03302445,0.70651054,-0.70633515,0.02903282],[-1,0,-1,0],[9E+09,9E+09,9E+09,9E+09,9E+09,9E+09]],[16.67,500,5000,1000],z1,Spindle \WObj:=Deburring;
		MoveL [[46.889,112.744,17.313],[0.03461177,0.70658837,-0.70625876,0.02708256],[-1,0,-1,0],[9E+09,9E+09,9E+09,9E+09,9E+09,9E+09]],[16.67,500,5000,1000],z1,Spindle \WObj:=Deburring;
		MoveL [[47.822,112.620,17.313],[0.03645880,0.70668746,-0.70616671,0.02433424],[-1,0,-1,0],[9E+09,9E+09,9E+09,9E+09,9E+09,9E+09]],[16.67,500,5000,1000],z1,Spindle \WObj:=Deburring;
		MoveL [[48.605,112.452,17.313],[0.03843428,0.70680808,-0.70606132,0.02055616],[-1,0,-1,0],[9E+09,9E+09,9E+09,9E+09,9E+09,9E+09]],[16.67,500,5000,1000],z1,Spindle \WObj:=Deburring;
		MoveL [[49.018,112.327,17.313],[0.03957779,0.70687059,-0.70599847,0.01826813],[-1,0,-1,0],[9E+09,9E+09,9E+09,9E+09,9E+09,9E+09]],[16.67,500,5000,1000],z1,Spindle \WObj:=Deburring;
		MoveL [[49.512,112.110,17.313],[0.04156894,0.70698183,-0.70588386,0.01329242],[-1,0,-1,0],[9E+09,9E+09,9E+09,9E+09,9E+09,9E+09]],[16.67,500,5000,1000],z1,Spindle \WObj:=Deburring;
		MoveL [[49.858,111.901,17.313],[0.04292705,0.70706553,-0.70580232,0.00766116],[-1,0,-1,0],[9E+09,9E+09,9E+09,9E+09,9E+09,9E+09]],[16.67,500,5000,1000],z1,Spindle \WObj:=Deburring;
		MoveL [[50.174,111.649,17.313],[0.04353448,0.70710350,-0.70576536,0.00215694],[-1,0,-1,0],[9E+09,9E+09,9E+09,9E+09,9E+09,9E+09]],[16.67,500,5000,1000],z1,Spindle \WObj:=Deburring;
		MoveL [[50.443,111.372,17.313],[0.04356951,0.70709828,-0.70576318,-0.00347112],[-1,0,-1,0],[9E+09,9E+09,9E+09,9E+09,9E+09,9E+09]],[16.67,500,5000,1000],z1,Spindle \WObj:=Deburring;
		MoveL [[50.734,110.959,17.313],[0.04219231,0.70701131,-0.70584655,-0.01163885],[-1,0,-1,0],[9E+09,9E+09,9E+09,9E+09,9E+09,9E+09]],[16.67,500,5000,1000],z1,Spindle \WObj:=Deburring;
		MoveL [[50.884,110.696,17.313],[0.04123080,0.70696589,-0.70590365,-0.01411685],[-1,0,-1,0],[9E+09,9E+09,9E+09,9E+09,9E+09,9E+09]],[16.67,500,5000,1000],z1,Spindle \WObj:=Deburring;
		MoveL [[51.091,110.198,17.313],[0.03929315,0.70685324,-0.70601414,-0.01893607],[-1,0,-1,0],[9E+09,9E+09,9E+09,9E+09,9E+09,9E+09]],[16.67,500,5000,1000],z1,Spindle \WObj:=Deburring;
		MoveL [[51.292,109.435,17.313],[0.03570394,0.70666491,-0.70620502,-0.02498812],[-1,0,-1,0],[9E+09,9E+09,9E+09,9E+09,9E+09,9E+09]],[16.67,500,5000,1000],z1,Spindle \WObj:=Deburring;
		MoveL [[51.423,108.631,17.313],[0.03380015,0.70656777,-0.70629862,-0.02760046],[-1,0,-1,0],[9E+09,9E+09,9E+09,9E+09,9E+09,9E+09]],[16.67,500,5000,1000],z1,Spindle \WObj:=Deburring;
		MoveL [[51.537,107.419,17.313],[0.03235416,0.70650146,-0.70636645,-0.02924592],[-1,0,-1,0],[9E+09,9E+09,9E+09,9E+09,9E+09,9E+09]],[16.67,500,5000,1000],z1,Spindle \WObj:=Deburring;
		MoveL [[51.629,105.313,17.313],[0.03155438,0.70646044,-0.70640218,-0.03023125],[-1,0,-1,0],[9E+09,9E+09,9E+09,9E+09,9E+09,9E+09]],[16.67,500,5000,1000],z1,Spindle \WObj:=Deburring;
		MoveL [[51.694,101.429,17.313],[0.03098738,0.70644601,-0.70642739,-0.03056411],[-1,0,-1,0],[9E+09,9E+09,9E+09,9E+09,9E+09,9E+09]],[16.67,500,5000,1000],z1,Spindle \WObj:=Deburring;
		MoveL [[51.708,97.775,17.313],[0.03098738,0.70644601,-0.70642739,-0.03056411],[-1,0,-1,0],[9E+09,9E+09,9E+09,9E+09,9E+09,9E+09]],[16.67,500,5000,1000],z1,Spindle \WObj:=Deburring;
		MoveL [[51.722,94.121,17.313],[0.03092991,0.70643988,-0.70642980,-0.03070790],[-1,0,-1,0],[9E+09,9E+09,9E+09,9E+09,9E+09,9E+09]],[16.67,500,5000,1000],z1,Spindle \WObj:=Deburring;
		MoveL [[51.737,90.467,17.313],[0.03090425,0.70643668,-0.70643086,-0.03078287],[-1,0,-1,0],[9E+09,9E+09,9E+09,9E+09,9E+09,9E+09]],[16.67,500,5000,1000],z1,Spindle \WObj:=Deburring;
		MoveL [[51.737,85.601,17.313],[0.03090425,0.70643668,-0.70643086,-0.03078287],[-1,0,-1,0],[9E+09,9E+09,9E+09,9E+09,9E+09,9E+09]],[16.67,500,5000,1000],z1,Spindle \WObj:=Deburring;
		MoveL [[51.737,80.735,17.313],[0.03090425,0.70643668,-0.70643086,-0.03078287],[-1,0,-1,0],[9E+09,9E+09,9E+09,9E+09,9E+09,9E+09]],[16.67,500,5000,1000],z1,Spindle \WObj:=Deburring;
		MoveL [[51.737,75.869,17.313],[0.03090425,0.70643668,-0.70643086,-0.03078287],[-1,0,-1,0],[9E+09,9E+09,9E+09,9E+09,9E+09,9E+09]],[16.67,500,5000,1000],z1,Spindle \WObj:=Deburring;
		MoveL [[51.737,71.002,17.313],[0.03090425,0.70643668,-0.70643086,-0.03078287],[-1,0,-1,0],[9E+09,9E+09,9E+09,9E+09,9E+09,9E+09]],[16.67,500,5000,1000],z1,Spindle \WObj:=Deburring;
		MoveL [[51.738,66.136,17.313],[0.03090425,0.70643668,-0.70643086,-0.03078287],[-1,0,-1,0],[9E+09,9E+09,9E+09,9E+09,9E+09,9E+09]],[16.67,500,5000,1000],z1,Spindle \WObj:=Deburring;
		MoveL [[51.738,61.270,17.313],[0.03090425,0.70643668,-0.70643086,-0.03078287],[-1,0,-1,0],[9E+09,9E+09,9E+09,9E+09,9E+09,9E+09]],[16.67,500,5000,1000],z1,Spindle \WObj:=Deburring;
		MoveL [[51.738,56.404,17.313],[0.03090425,0.70643668,-0.70643086,-0.03078287],[-1,0,-1,0],[9E+09,9E+09,9E+09,9E+09,9E+09,9E+09]],[16.67,500,5000,1000],z1,Spindle \WObj:=Deburring;
		MoveL [[51.738,51.538,17.313],[0.03090425,0.70643668,-0.70643086,-0.03078287],[-1,0,-1,0],[9E+09,9E+09,9E+09,9E+09,9E+09,9E+09]],[16.67,500,5000,1000],z1,Spindle \WObj:=Deburring;
		MoveL [[51.739,46.672,17.313],[0.03090425,0.70643668,-0.70643086,-0.03078287],[-1,0,-1,0],[9E+09,9E+09,9E+09,9E+09,9E+09,9E+09]],[16.67,500,5000,1000],z1,Spindle \WObj:=Deburring;
		MoveL [[51.739,41.806,17.313],[0.03090425,0.70643668,-0.70643086,-0.03078287],[-1,0,-1,0],[9E+09,9E+09,9E+09,9E+09,9E+09,9E+09]],[16.67,500,5000,1000],z1,Spindle \WObj:=Deburring;
		MoveL [[51.739,36.939,17.313],[0.03090425,0.70643668,-0.70643086,-0.03078287],[-1,0,-1,0],[9E+09,9E+09,9E+09,9E+09,9E+09,9E+09]],[16.67,500,5000,1000],z1,Spindle \WObj:=Deburring;
		MoveL [[51.739,32.073,17.313],[0.03090425,0.70643668,-0.70643086,-0.03078287],[-1,0,-1,0],[9E+09,9E+09,9E+09,9E+09,9E+09,9E+09]],[16.67,500,5000,1000],z1,Spindle \WObj:=Deburring;
		MoveL [[51.739,27.207,17.313],[0.03090425,0.70643668,-0.70643086,-0.03078287],[-1,0,-1,0],[9E+09,9E+09,9E+09,9E+09,9E+09,9E+09]],[16.67,500,5000,1000],z1,Spindle \WObj:=Deburring;
		MoveL [[51.740,22.341,17.313],[0.03090425,0.70643668,-0.70643086,-0.03078287],[-1,0,-1,0],[9E+09,9E+09,9E+09,9E+09,9E+09,9E+09]],[16.67,500,5000,1000],z1,Spindle \WObj:=Deburring;
		MoveL [[51.740,17.475,17.313],[0.03090425,0.70643668,-0.70643086,-0.03078287],[-1,0,-1,0],[9E+09,9E+09,9E+09,9E+09,9E+09,9E+09]],[16.67,500,5000,1000],z1,Spindle \WObj:=Deburring;
		MoveL [[51.740,12.608,17.313],[0.03090425,0.70643668,-0.70643086,-0.03078287],[-1,0,-1,0],[9E+09,9E+09,9E+09,9E+09,9E+09,9E+09]],[16.67,500,5000,1000],z1,Spindle \WObj:=Deburring;
		MoveL [[51.740,7.742,17.313],[0.03090425,0.70643668,-0.70643086,-0.03078287],[-1,0,-1,0],[9E+09,9E+09,9E+09,9E+09,9E+09,9E+09]],[16.67,500,5000,1000],z1,Spindle \WObj:=Deburring;
		MoveL [[51.740,2.876,17.313],[0.03090425,0.70643668,-0.70643086,-0.03078287],[-1,0,-1,0],[9E+09,9E+09,9E+09,9E+09,9E+09,9E+09]],[16.67,500,5000,1000],z1,Spindle \WObj:=Deburring;
		MoveL [[51.741,-1.990,17.313],[0.03090425,0.70643668,-0.70643086,-0.03078287],[-1,0,-1,0],[9E+09,9E+09,9E+09,9E+09,9E+09,9E+09]],[16.67,500,5000,1000],z1,Spindle \WObj:=Deburring;
		MoveL [[51.741,-6.856,17.313],[0.03090425,0.70643668,-0.70643086,-0.03078287],[-1,0,-1,0],[9E+09,9E+09,9E+09,9E+09,9E+09,9E+09]],[16.67,500,5000,1000],z1,Spindle \WObj:=Deburring;
		MoveL [[51.741,-11.722,17.313],[0.03090425,0.70643668,-0.70643086,-0.03078287],[-1,0,-1,0],[9E+09,9E+09,9E+09,9E+09,9E+09,9E+09]],[16.67,500,5000,1000],z1,Spindle \WObj:=Deburring;
		MoveL [[51.741,-16.588,17.313],[0.03090425,0.70643668,-0.70643086,-0.03078287],[-1,0,-1,0],[9E+09,9E+09,9E+09,9E+09,9E+09,9E+09]],[16.67,500,5000,1000],z1,Spindle \WObj:=Deburring;
		MoveL [[51.742,-21.455,17.313],[0.03090425,0.70643668,-0.70643086,-0.03078287],[-1,0,-1,0],[9E+09,9E+09,9E+09,9E+09,9E+09,9E+09]],[16.67,500,5000,1000],z1,Spindle \WObj:=Deburring;
		MoveL [[51.742,-26.321,17.313],[0.03090425,0.70643668,-0.70643086,-0.03078287],[-1,0,-1,0],[9E+09,9E+09,9E+09,9E+09,9E+09,9E+09]],[16.67,500,5000,1000],z1,Spindle \WObj:=Deburring;
		MoveL [[51.742,-31.187,17.313],[0.03090425,0.70643668,-0.70643086,-0.03078287],[-1,0,-1,0],[9E+09,9E+09,9E+09,9E+09,9E+09,9E+09]],[16.67,500,5000,1000],z1,Spindle \WObj:=Deburring;
		MoveL [[51.742,-36.053,17.313],[0.03090425,0.70643668,-0.70643086,-0.03078287],[-1,0,-1,0],[9E+09,9E+09,9E+09,9E+09,9E+09,9E+09]],[16.67,500,5000,1000],z1,Spindle \WObj:=Deburring;
		MoveL [[51.742,-40.919,17.313],[0.03090425,0.70643668,-0.70643086,-0.03078287],[-1,0,-1,0],[9E+09,9E+09,9E+09,9E+09,9E+09,9E+09]],[16.67,500,5000,1000],z1,Spindle \WObj:=Deburring;
		MoveL [[51.743,-45.785,17.313],[0.03090425,0.70643668,-0.70643086,-0.03078287],[-1,0,-1,0],[9E+09,9E+09,9E+09,9E+09,9E+09,9E+09]],[16.67,500,5000,1000],z1,Spindle \WObj:=Deburring;
		MoveL [[51.743,-50.651,17.313],[0.03090425,0.70643668,-0.70643086,-0.03078287],[-1,0,-1,0],[9E+09,9E+09,9E+09,9E+09,9E+09,9E+09]],[16.67,500,5000,1000],z1,Spindle \WObj:=Deburring;
		MoveL [[51.743,-55.518,17.313],[0.03090425,0.70643668,-0.70643086,-0.03078287],[-1,0,-1,0],[9E+09,9E+09,9E+09,9E+09,9E+09,9E+09]],[16.67,500,5000,1000],z1,Spindle \WObj:=Deburring;
		MoveL [[51.743,-60.384,17.313],[0.03090425,0.70643668,-0.70643086,-0.03078287],[-1,0,-1,0],[9E+09,9E+09,9E+09,9E+09,9E+09,9E+09]],[16.67,500,5000,1000],z1,Spindle \WObj:=Deburring;
		MoveL [[51.743,-65.250,17.313],[0.03090425,0.70643668,-0.70643086,-0.03078287],[-1,0,-1,0],[9E+09,9E+09,9E+09,9E+09,9E+09,9E+09]],[16.67,500,5000,1000],z1,Spindle \WObj:=Deburring;
		MoveL [[51.744,-70.116,17.313],[0.03090425,0.70643668,-0.70643086,-0.03078287],[-1,0,-1,0],[9E+09,9E+09,9E+09,9E+09,9E+09,9E+09]],[16.67,500,5000,1000],z1,Spindle \WObj:=Deburring;
		MoveL [[51.744,-74.982,17.313],[0.03088059,0.70643524,-0.70643230,-0.03080654],[-1,0,-1,0],[9E+09,9E+09,9E+09,9E+09,9E+09,9E+09]],[16.67,500,5000,1000],z1,Spindle \WObj:=Deburring;
		MoveL [[51.740,-79.353,17.313],[0.03088059,0.70643524,-0.70643230,-0.03080654],[-1,0,-1,0],[9E+09,9E+09,9E+09,9E+09,9E+09,9E+09]],[16.67,500,5000,1000],z1,Spindle \WObj:=Deburring;
		MoveL [[51.736,-83.725,17.313],[0.03081437,0.70643196,-0.70643505,-0.03088508],[-1,0,-1,0],[9E+09,9E+09,9E+09,9E+09,9E+09,9E+09]],[16.67,500,5000,1000],z1,Spindle \WObj:=Deburring;
		MoveL [[51.732,-88.096,17.313],[0.03078435,0.70643018,-0.70643628,-0.03092744],[-1,0,-1,0],[9E+09,9E+09,9E+09,9E+09,9E+09,9E+09]],[16.67,500,5000,1000],z1,Spindle \WObj:=Deburring;
		MoveL [[51.728,-92.467,17.313],[0.03075432,0.70642840,-0.70643751,-0.03096979],[-1,0,-1,0],[9E+09,9E+09,9E+09,9E+09,9E+09,9E+09]],[16.67,500,5000,1000],z1,Spindle \WObj:=Deburring;
		MoveL [[51.724,-96.838,17.313],[0.03072429,0.70642662,-0.70643874,-0.03101215],[-1,0,-1,0],[9E+09,9E+09,9E+09,9E+09,9E+09,9E+09]],[16.67,500,5000,1000],z1,Spindle \WObj:=Deburring;
		MoveL [[51.699,-100.136,17.313],[0.03045872,0.70641650,-0.70645029,-0.03124070],[-1,0,-1,0],[9E+09,9E+09,9E+09,9E+09,9E+09,9E+09]],[16.67,500,5000,1000],z1,Spindle \WObj:=Deburring;
		MoveL [[51.673,-103.433,17.313],[0.03019928,0.70640602,-0.70646149,-0.03147539],[-1,0,-1,0],[9E+09,9E+09,9E+09,9E+09,9E+09,9E+09]],[16.67,500,5000,1000],z1,Spindle \WObj:=Deburring;
		MoveL [[51.602,-106.266,17.313],[0.02912333,0.70636472,-0.70650660,-0.03239037],[-1,0,-1,0],[9E+09,9E+09,9E+09,9E+09,9E+09,9E+09]],[16.67,500,5000,1000],z1,Spindle \WObj:=Deburring;
		MoveL [[51.507,-107.903,17.313],[0.02743446,0.70629397,-0.70657449,-0.03389192],[-1,0,-1,0],[9E+09,9E+09,9E+09,9E+09,9E+09,9E+09]],[16.67,500,5000,1000],z1,Spindle \WObj:=Deburring;
		MoveL [[51.384,-108.970,17.313],[0.02477336,0.70620085,-0.70667265,-0.03578260],[-1,0,-1,0],[9E+09,9E+09,9E+09,9E+09,9E+09,9E+09]],[16.67,500,5000,1000],z1,Spindle \WObj:=Deburring;
		MoveL [[51.229,-109.756,17.313],[0.02151229,0.70608233,-0.70677964,-0.03804610],[-1,0,-1,0],[9E+09,9E+09,9E+09,9E+09,9E+09,9E+09]],[16.67,500,5000,1000],z1,Spindle \WObj:=Deburring;
		MoveL [[51.073,-110.272,17.313],[0.01731601,0.70596317,-0.70689454,-0.04020286],[-1,0,-1,0],[9E+09,9E+09,9E+09,9E+09,9E+09,9E+09]],[16.67,500,5000,1000],z1,Spindle \WObj:=Deburring;
		MoveL [[50.914,-110.673,17.313],[0.01478322,0.70592022,-0.70695205,-0.04094989],[-1,0,-1,0],[9E+09,9E+09,9E+09,9E+09,9E+09,9E+09]],[16.67,500,5000,1000],z1,Spindle \WObj:=Deburring;
		MoveL [[50.670,-111.094,17.313],[0.00739238,0.70579861,-0.70706807,-0.04299320],[-1,0,-1,0],[9E+09,9E+09,9E+09,9E+09,9E+09,9E+09]],[16.67,500,5000,1000],z1,Spindle \WObj:=Deburring;
		MoveL [[50.426,-111.415,17.313],[0.00181340,0.70576709,-0.70710432,-0.04350874],[-1,0,-1,0],[9E+09,9E+09,9E+09,9E+09,9E+09,9E+09]],[16.67,500,5000,1000],z1,Spindle \WObj:=Deburring;
		MoveL [[50.221,-111.638,17.313],[0.00103582,-0.70576468,0.70710571,0.04355064],[-1,0,-1,0],[9E+09,9E+09,9E+09,9E+09,9E+09,9E+09]],[16.67,500,5000,1000],z1,Spindle \WObj:=Deburring;
		MoveL [[49.909,-111.896,17.313],[0.00685774,-0.70580554,0.70707355,0.04287768],[-1,0,-1,0],[9E+09,9E+09,9E+09,9E+09,9E+09,9E+09]],[16.67,500,5000,1000],z1,Spindle \WObj:=Deburring;
		MoveL [[49.567,-112.111,17.313],[0.01249303,-0.70588296,0.70699642,0.04158395],[-1,0,-1,0],[9E+09,9E+09,9E+09,9E+09,9E+09,9E+09]],[16.67,500,5000,1000],z1,Spindle \WObj:=Deburring;
		MoveL [[49.076,-112.333,17.313],[0.01764733,-0.70598035,0.70688680,0.03989185],[-1,0,-1,0],[9E+09,9E+09,9E+09,9E+09,9E+09,9E+09]],[16.67,500,5000,1000],z1,Spindle \WObj:=Deburring;
		MoveL [[48.449,-112.521,17.313],[0.02374797,-0.70616017,0.70670802,0.03657358],[-1,0,-1,0],[9E+09,9E+09,9E+09,9E+09,9E+09,9E+09]],[16.67,500,5000,1000],z1,Spindle \WObj:=Deburring;
		MoveL [[47.652,-112.680,17.313],[0.02672742,-0.70626857,0.70660160,0.03441697],[-1,0,-1,0],[9E+09,9E+09,9E+09,9E+09,9E+09,9E+09]],[16.67,500,5000,1000],z1,Spindle \WObj:=Deburring;
		MoveL [[46.578,-112.808,17.313],[0.02874819,-0.70634370,0.70652230,0.03283837],[-1,0,-1,0],[9E+09,9E+09,9E+09,9E+09,9E+09,9E+09]],[16.67,500,5000,1000],z1,Spindle \WObj:=Deburring;
		MoveL [[44.997,-112.903,17.313],[0.03004715,-0.70639610,0.70646761,0.03170533],[-1,0,-1,0],[9E+09,9E+09,9E+09,9E+09,9E+09,9E+09]],[16.67,500,5000,1000],z1,Spindle \WObj:=Deburring;
		MoveL [[42.459,-112.960,17.313],[0.03067067,-0.70643084,0.70644159,0.03090402],[-1,0,-1,0],[9E+09,9E+09,9E+09,9E+09,9E+09,9E+09]],[16.67,500,5000,1000],z1,Spindle \WObj:=Deburring;
		MoveL [[37.896,-112.971,17.313],[0.03081561,-0.70643007,0.70643508,0.03092614],[-1,0,-1,0],[9E+09,9E+09,9E+09,9E+09,9E+09,9E+09]],[16.67,500,5000,1000],z1,Spindle \WObj:=Deburring;
		MoveL [[33.332,-112.982,17.313],[0.03096662,-0.70642962,0.70642823,0.03094207],[-1,0,-1,0],[9E+09,9E+09,9E+09,9E+09,9E+09,9E+09]],[16.67,500,5000,1000],z1,Spindle \WObj:=Deburring;
		MoveL [[28.430,-112.980,17.313],[0.03096662,-0.70642962,0.70642823,0.03094207],[-1,0,-1,0],[9E+09,9E+09,9E+09,9E+09,9E+09,9E+09]],[16.67,500,5000,1000],z1,Spindle \WObj:=Deburring;
		MoveL [[23.528,-112.978,17.313],[0.03096662,-0.70642962,0.70642823,0.03094207],[-1,0,-1,0],[9E+09,9E+09,9E+09,9E+09,9E+09,9E+09]],[16.67,500,5000,1000],z1,Spindle \WObj:=Deburring;
		MoveL [[18.625,-112.976,17.313],[0.03096662,-0.70642962,0.70642823,0.03094207],[-1,0,-1,0],[9E+09,9E+09,9E+09,9E+09,9E+09,9E+09]],[16.67,500,5000,1000],z1,Spindle \WObj:=Deburring;
		MoveL [[13.723,-112.974,17.313],[0.03096662,-0.70642962,0.70642823,0.03094207],[-1,0,-1,0],[9E+09,9E+09,9E+09,9E+09,9E+09,9E+09]],[16.67,500,5000,1000],z1,Spindle \WObj:=Deburring;
		MoveL [[8.821,-112.972,17.313],[0.03096662,-0.70642962,0.70642823,0.03094207],[-1,0,-1,0],[9E+09,9E+09,9E+09,9E+09,9E+09,9E+09]],[16.67,500,5000,1000],z1,Spindle \WObj:=Deburring;
		MoveL [[3.919,-112.970,17.313],[0.03096662,-0.70642962,0.70642823,0.03094207],[-1,0,-1,0],[9E+09,9E+09,9E+09,9E+09,9E+09,9E+09]],[16.67,500,5000,1000],z1,Spindle \WObj:=Deburring;
		MoveL [[-0.983,-112.968,17.313],[0.03088878,-0.70642687,0.70643188,0.03099932],[0,-1,0,0],[9E+09,9E+09,9E+09,9E+09,9E+09,9E+09]],[16.67,500,5000,1000],z1,Spindle \WObj:=Deburring;
		MoveL [[-5.886,-112.965,17.313],[0.03088117,-0.70642659,0.70643229,0.03100398],[0,-1,0,0],[9E+09,9E+09,9E+09,9E+09,9E+09,9E+09]],[16.67,500,5000,1000],z1,Spindle \WObj:=Deburring;
		MoveL [[-10.788,-112.963,17.313],[0.03086745,-0.70642658,0.70643243,0.03101486],[0,-1,0,0],[9E+09,9E+09,9E+09,9E+09,9E+09,9E+09]],[16.67,500,5000,1000],z1,Spindle \WObj:=Deburring;
		MoveL [[-15.690,-112.961,17.313],[0.03085986,-0.70642568,0.70643345,0.03101949],[0,-1,0,0],[9E+09,9E+09,9E+09,9E+09,9E+09,9E+09]],[16.67,500,5000,1000],z1,Spindle \WObj:=Deburring;
		MoveL [[-20.592,-112.959,17.313],[0.03084607,-0.70642566,0.70643359,0.03103032],[0,-1,0,0],[9E+09,9E+09,9E+09,9E+09,9E+09,9E+09]],[16.67,500,5000,1000],z1,Spindle \WObj:=Deburring;
		MoveL [[-25.494,-112.957,17.313],[0.03083846,-0.70642538,0.70643400,0.03103497],[0,-1,0,0],[9E+09,9E+09,9E+09,9E+09,9E+09,9E+09]],[16.67,500,5000,1000],z1,Spindle \WObj:=Deburring;
		MoveL [[-30.396,-112.955,17.313],[0.03082470,-0.70642475,0.70643476,0.03104577],[0,-1,0,0],[9E+09,9E+09,9E+09,9E+09,9E+09,9E+09]],[16.67,500,5000,1000],z1,Spindle \WObj:=Deburring;
		MoveL [[-35.299,-112.953,17.313],[0.03081709,-0.70642447,0.70643517,0.03105043],[0,-1,0,0],[9E+09,9E+09,9E+09,9E+09,9E+09,9E+09]],[16.67,500,5000,1000],z1,Spindle \WObj:=Deburring;
		MoveL [[-39.452,-112.951,17.313],[0.03103952,-0.70643996,0.70642545,0.03069558],[0,-1,0,0],[9E+09,9E+09,9E+09,9E+09,9E+09,9E+09]],[16.67,500,5000,1000],z1,Spindle \WObj:=Deburring;
		MoveL [[-43.128,-112.925,17.313],[0.03085198,-0.70647033,0.70643351,0.02999207],[0,-1,0,0],[9E+09,9E+09,9E+09,9E+09,9E+09,9E+09]],[16.67,500,5000,1000],z1,Spindle \WObj:=Deburring;
		MoveL [[-44.856,-112.889,17.313],[0.03187801,-0.70650169,0.70638825,0.02923697],[0,-1,0,0],[9E+09,9E+09,9E+09,9E+09,9E+09,9E+09]],[16.67,500,5000,1000],z1,Spindle \WObj:=Deburring;
		MoveL [[-46.221,-112.819,17.313],[0.03358530,-0.70656287,0.70630886,0.02772613],[0,-1,0,0],[9E+09,9E+09,9E+09,9E+09,9E+09,9E+09]],[16.67,500,5000,1000],z1,Spindle \WObj:=Deburring;
		MoveL [[-47.420,-112.699,17.313],[0.03531810,-0.70664573,0.70622431,0.02552760],[0,-1,0,0],[9E+09,9E+09,9E+09,9E+09,9E+09,9E+09]],[16.67,500,5000,1000],z1,Spindle \WObj:=Deburring;
		MoveL [[-48.198,-112.565,17.313],[0.03740543,-0.70674508,0.70611634,0.02262593],[0,-1,0,0],[9E+09,9E+09,9E+09,9E+09,9E+09,9E+09]],[16.67,500,5000,1000],z1,Spindle \WObj:=Deburring;
		MoveL [[-48.846,-112.395,17.313],[0.03954608,-0.70686434,0.70599995,0.01851975],[0,-1,0,0],[9E+09,9E+09,9E+09,9E+09,9E+09,9E+09]],[16.67,500,5000,1000],z1,Spindle \WObj:=Deburring;
		MoveL [[-49.342,-112.203,17.313],[0.04136766,-0.70697268,0.70589573,0.01376828],[0,-1,0,0],[9E+09,9E+09,9E+09,9E+09,9E+09,9E+09]],[16.67,500,5000,1000],z1,Spindle \WObj:=Deburring;
		MoveL [[-49.698,-112.012,17.313],[0.04284762,-0.70705174,0.70580717,0.00884094],[0,-1,0,0],[9E+09,9E+09,9E+09,9E+09,9E+09,9E+09]],[16.67,500,5000,1000],z1,Spindle \WObj:=Deburring;
		MoveL [[-50.028,-111.781,17.313],[0.04362403,-0.70709841,0.70575944,0.00352061],[0,-1,0,0],[9E+09,9E+09,9E+09,9E+09,9E+09,9E+09]],[16.67,500,5000,1000],z1,Spindle \WObj:=Deburring;
		MoveL [[-50.259,-111.584,17.313],[0.04365796,-0.70710717,0.70575726,0.00034053],[0,-1,0,0],[9E+09,9E+09,9E+09,9E+09,9E+09,9E+09]],[16.67,500,5000,1000],z1,Spindle \WObj:=Deburring;
		MoveL [[-50.529,-111.283,17.313],[0.04320163,-0.70708537,0.70578575,-0.00551219],[0,-1,0,0],[9E+09,9E+09,9E+09,9E+09,9E+09,9E+09]],[16.67,500,5000,1000],z1,Spindle \WObj:=Deburring;
		MoveL [[-50.803,-110.859,17.313],[0.04155807,-0.70698427,0.70588483,-0.01314399],[0,-1,0,0],[9E+09,9E+09,9E+09,9E+09,9E+09,9E+09]],[16.67,500,5000,1000],z1,Spindle \WObj:=Deburring;
		MoveL [[-50.981,-110.489,17.313],[0.03976293,-0.70687998,0.70598791,-0.01790712],[0,-1,0,0],[9E+09,9E+09,9E+09,9E+09,9E+09,9E+09]],[16.67,500,5000,1000],z1,Spindle \WObj:=Deburring;
		MoveL [[-51.135,-110.086,17.313],[0.03867973,-0.70682049,0.70604801,-0.02012154],[0,-1,0,0],[9E+09,9E+09,9E+09,9E+09,9E+09,9E+09]],[16.67,500,5000,1000],z1,Spindle \WObj:=Deburring;
		MoveL [[-51.320,-109.325,17.313],[0.03555882,-0.70665494,0.70621186,-0.02528187],[0,-1,0,0],[9E+09,9E+09,9E+09,9E+09,9E+09,9E+09]],[16.67,500,5000,1000],z1,Spindle \WObj:=Deburring;
		MoveL [[-51.411,-108.786,17.313],[0.03465069,-0.70660993,0.70625734,-0.02650120],[0,-1,0,0],[9E+09,9E+09,9E+09,9E+09,9E+09,9E+09]],[16.67,500,5000,1000],z1,Spindle \WObj:=Deburring;
		MoveL [[-51.537,-107.460,17.313],[0.03240548,-0.70649726,0.70636378,-0.02935491],[0,-1,0,0],[9E+09,9E+09,9E+09,9E+09,9E+09,9E+09]],[16.67,500,5000,1000],z1,Spindle \WObj:=Deburring;
		MoveL [[-51.631,-105.330,17.313],[0.03136553,-0.70646205,0.70641092,-0.03018586],[0,-1,0,0],[9E+09,9E+09,9E+09,9E+09,9E+09,9E+09]],[16.67,500,5000,1000],z1,Spindle \WObj:=Deburring;
		MoveL [[-51.697,-101.334,17.313],[0.03097875,-0.70644083,0.70642776,-0.03068371],[0,-1,0,0],[9E+09,9E+09,9E+09,9E+09,9E+09,9E+09]],[16.67,500,5000,1000],z1,Spindle \WObj:=Deburring;
		MoveL [[-51.711,-97.477,17.313],[0.03097875,-0.70644083,0.70642776,-0.03068371],[0,-1,0,0],[9E+09,9E+09,9E+09,9E+09,9E+09,9E+09]],[16.67,500,5000,1000],z1,Spindle \WObj:=Deburring;
		MoveL [[-51.725,-93.620,17.313],[0.03083290,-0.70643856,0.70643436,-0.03073093],[0,-1,0,0],[9E+09,9E+09,9E+09,9E+09,9E+09,9E+09]],[16.67,500,5000,1000],z1,Spindle \WObj:=Deburring;
		MoveL [[-51.739,-89.762,17.313],[0.03075997,-0.70643742,0.70643765,-0.03075455],[0,-1,0,0],[9E+09,9E+09,9E+09,9E+09,9E+09,9E+09]],[16.67,500,5000,1000],z1,Spindle \WObj:=Deburring;
		MoveL [[-51.740,-86.623,17.313],[0.05960304,-0.70710237,0.70459039,-0.00247176],[0,-1,0,0],[9E+09,9E+09,9E+09,9E+09,9E+09,9E+09]],[16.67,500,5000,1000],z1,Spindle \WObj:=Deburring;
		MoveL [[-51.740,-83.483,17.313],[0.08834616,-0.70663544,0.70156602,0.02581523],[0,-1,0,0],[9E+09,9E+09,9E+09,9E+09,9E+09,9E+09]],[16.67,500,5000,1000],z1,Spindle \WObj:=Deburring;
		MoveL [[-51.740,-80.343,17.313],[0.11694896,-0.70503799,0.69736838,0.05405289],[0,-1,0,0],[9E+09,9E+09,9E+09,9E+09,9E+09,9E+09]],[16.67,500,5000,1000],z1,Spindle \WObj:=Deburring;
		MoveL [[-51.752,-80.314,17.312],[0.11694896,-0.70503799,0.69736838,0.05405289],[0,-1,0,0],[9E+09,9E+09,9E+09,9E+09,9E+09,9E+09]],[16.67,500,5000,1000],z1,Spindle \WObj:=Deburring;
		MoveL [[-51.780,-80.303,17.309],[0.11694896,-0.70503799,0.69736838,0.05405289],[0,-1,0,0],[9E+09,9E+09,9E+09,9E+09,9E+09,9E+09]],[16.67,500,5000,1000],z1,Spindle \WObj:=Deburring;
		MoveL [[-51.805,-80.283,17.307],[0.11694896,-0.70503799,0.69736838,0.05405289],[0,-1,0,0],[9E+09,9E+09,9E+09,9E+09,9E+09,9E+09]],[16.67,500,5000,1000],z1,Spindle \WObj:=Deburring;
		MoveL [[-51.832,-80.267,17.319],[0.11694896,-0.70503799,0.69736838,0.05405289],[0,-1,0,0],[9E+09,9E+09,9E+09,9E+09,9E+09,9E+09]],[16.67,500,5000,1000],z1,Spindle \WObj:=Deburring;
		MoveL [[-51.845,-80.266,17.349],[0.11694896,-0.70503799,0.69736838,0.05405289],[0,-1,0,0],[9E+09,9E+09,9E+09,9E+09,9E+09,9E+09]],[16.67,500,5000,1000],z1,Spindle \WObj:=Deburring;
		MoveL [[-52.286,-81.484,22.248],[0.11694896,-0.70503799,0.69736838,0.05405289],[0,-1,0,0],[9E+09,9E+09,9E+09,9E+09,9E+09,9E+09]],v1000,z1,Spindle \WObj:=Deburring;
		MoveL [[-52.286,-81.484,86.000],[0.11694896,-0.70503799,0.69736838,0.05405289],[0,-1,0,0],[9E+09,9E+09,9E+09,9E+09,9E+09,9E+09]],v1000,z1,Spindle \WObj:=Deburring;
		MoveL [[-52.286,-81.484,86.000],[0.11694896,-0.70503799,0.69736838,0.05405289],[0,-1,0,0],[9E+09,9E+09,9E+09,9E+09,9E+09,9E+09]],v1000,z1,Spindle \WObj:=Deburring;
		Spindle 0;
	ENDPROC

	PROC PickStation()
		ConfJ \On;
		ConfL \Off;
		PartStation := [FALSE, TRUE, "", [[0,0,0],[1,0,0,0]],[[620.000,0.000,396.884],[0.70710678,0.00000000,0.00000000,-0.70710678]]];
		SuctionCup := [TRUE,[[-94.709,0.000,259.352],[0.00000000,0.00000000,0.00000000,1.00000000]],[1,[0,0,20],[1,0,0,0],0,0,0.005]];
		MoveAbsJ [[9.440500,34.191600,-49.511700,0.000000,105.320000,99.440500],[9E+09,9E+09,9E+09,9E+09,9E+09,9E+09]],v1000,z1,SuctionCup \WObj:=PartStation;
		MoveL [[-16.111,46.392,100.500],[0.00000000,1.00000000,0.00000000,-0.00000000],[0,2,-1,1],[9E+09,9E+09,9E+09,9E+09,9E+09,9E+09]],v1000,z1,SuctionCup \WObj:=PartStation;
		! Attach to Suction Cup
		WaitTime 0.500;
		MoveL [[-16.111,46.485,191.000],[0.00000000,1.00000000,0.00000000,-0.00000000],[0,0,1,0],[9E+09,9E+09,9E+09,9E+09,9E+09,9E+09]],v1000,z1,SuctionCup \WObj:=PartStation;
	ENDPROC

	PROC DropOut1()
		ConfJ \On;
		ConfL \Off;
		SuctionCup := [TRUE,[[-94.709,0.000,259.352],[0.00000000,0.00000000,0.00000000,1.00000000]],[1,[0,0,20],[1,0,0,0],0,0,0.005]];
		MoveAbsJ [[-66.056500,21.575200,36.080800,0.000000,32.344000,-66.056500],[9E+09,9E+09,9E+09,9E+09,9E+09,9E+09]],v1000,z1,SuctionCup \WObj:=Out;
		MoveL [[-16.111,46.392,30.000],[0.00000000,1.00000000,0.00000000,-0.00000000],[-1,0,-1,0],[9E+09,9E+09,9E+09,9E+09,9E+09,9E+09]],v1000,z1,SuctionCup \WObj:=Out;
		! Detach from Suction Cup
		WaitTime 0.500;
		MoveL [[-16.111,46.485,105.701],[0.00000000,1.00000000,0.00000000,-0.00000000],[-1,0,-1,0],[9E+09,9E+09,9E+09,9E+09,9E+09,9E+09]],v1000,z1,SuctionCup \WObj:=Out;
	ENDPROC

	PROC PickIn2()
		ConfJ \On;
		ConfL \Off;
		In := [FALSE, TRUE, "", [[0,0,0],[1,0,0,0]],[[290.000,450.000,10.000],[1.00000000,0.00000000,0.00000000,0.00000000]]];
		SuctionCup := [TRUE,[[-94.709,0.000,259.352],[0.00000000,0.00000000,0.00000000,1.00000000]],[1,[0,0,20],[1,0,0,0],0,0,0.005]];
		MoveAbsJ [[70.152800,32.938500,23.515600,0.000000,33.545900,70.152800],[9E+09,9E+09,9E+09,9E+09,9E+09,9E+09]],v1000,z1,SuctionCup \WObj:=In;
		MoveL [[-16.111,46.392,40.000],[0.00000000,1.00000000,0.00000000,-0.00000000],[0,2,-2,1],[9E+09,9E+09,9E+09,9E+09,9E+09,9E+09]],v1000,z1,SuctionCup \WObj:=In;
		! Attach to Suction Cup
		WaitTime 0.500;
		MoveL [[-16.087,46.472,70.960],[0.00000000,1.00000000,0.00000000,-0.00000000],[0,0,0,0],[9E+09,9E+09,9E+09,9E+09,9E+09,9E+09]],v1000,z1,SuctionCup \WObj:=In;
	ENDPROC

	PROC DropOut2()
		ConfJ \On;
		ConfL \Off;
		Out := [FALSE, TRUE, "", [[0,0,0],[1,0,0,0]],[[290.000,-450.000,10.000],[1.00000000,0.00000000,0.00000000,0.00000000]]];
		SuctionCup := [TRUE,[[-94.709,0.000,259.352],[0.00000000,0.00000000,0.00000000,1.00000000]],[1,[0,0,20],[1,0,0,0],0,0,0.005]];
		MoveAbsJ [[-66.056500,21.575200,36.080800,0.000000,32.344000,-66.056500],[9E+09,9E+09,9E+09,9E+09,9E+09,9E+09]],v1000,z1,SuctionCup \WObj:=Out;
		MoveL [[-16.111,46.392,35.000],[0.00000000,1.00000000,0.00000000,-0.00000000],[-1,0,-1,0],[9E+09,9E+09,9E+09,9E+09,9E+09,9E+09]],v1000,z1,SuctionCup \WObj:=Out;
		! Detach from Suction Cup
		WaitTime 0.500;
		MoveL [[-16.111,46.485,105.701],[0.00000000,1.00000000,0.00000000,-0.00000000],[-1,0,-1,0],[9E+09,9E+09,9E+09,9E+09,9E+09,9E+09]],v1000,z1,SuctionCup \WObj:=Out;
	ENDPROC

	PROC PickIn3()
		ConfJ \On;
		ConfL \Off;
		In := [FALSE, TRUE, "", [[0,0,0],[1,0,0,0]],[[290.000,450.000,10.000],[1.00000000,0.00000000,0.00000000,0.00000000]]];
		SuctionCup := [TRUE,[[-94.709,0.000,259.352],[0.00000000,0.00000000,0.00000000,1.00000000]],[1,[0,0,20],[1,0,0,0],0,0,0.005]];
		MoveAbsJ [[70.152800,32.938500,23.515600,0.000000,33.545900,70.152800],[9E+09,9E+09,9E+09,9E+09,9E+09,9E+09]],v1000,z1,SuctionCup \WObj:=In;
		MoveL [[-16.111,46.392,35.000],[0.00000000,1.00000000,0.00000000,-0.00000000],[0,2,-2,1],[9E+09,9E+09,9E+09,9E+09,9E+09,9E+09]],v1000,z1,SuctionCup \WObj:=In;
		! Attach to Suction Cup
		WaitTime 0.500;
		MoveL [[-16.087,46.472,70.960],[0.00000000,1.00000000,0.00000000,-0.00000000],[0,0,0,0],[9E+09,9E+09,9E+09,9E+09,9E+09,9E+09]],v1000,z1,SuctionCup \WObj:=In;
	ENDPROC

	PROC DropOut3()
		ConfJ \On;
		ConfL \Off;
		Out := [FALSE, TRUE, "", [[0,0,0],[1,0,0,0]],[[290.000,-450.000,10.000],[1.00000000,0.00000000,0.00000000,0.00000000]]];
		SuctionCup := [TRUE,[[-94.709,0.000,259.352],[0.00000000,0.00000000,0.00000000,1.00000000]],[1,[0,0,20],[1,0,0,0],0,0,0.005]];
		MoveAbsJ [[-66.056500,21.575200,36.080800,0.000000,32.344000,-66.056500],[9E+09,9E+09,9E+09,9E+09,9E+09,9E+09]],v1000,z1,SuctionCup \WObj:=Out;
		MoveL [[-16.111,46.392,40.000],[0.00000000,1.00000000,0.00000000,-0.00000000],[-1,0,-1,0],[9E+09,9E+09,9E+09,9E+09,9E+09,9E+09]],v1000,z1,SuctionCup \WObj:=Out;
		! Detach from Suction Cup
		WaitTime 0.500;
		MoveL [[-16.111,46.485,105.701],[0.00000000,1.00000000,0.00000000,-0.00000000],[-1,0,-1,0],[9E+09,9E+09,9E+09,9E+09,9E+09,9E+09]],v1000,z1,SuctionCup \WObj:=Out;
	ENDPROC

	PROC PickIn4()
		ConfJ \On;
		ConfL \Off;
		In := [FALSE, TRUE, "", [[0,0,0],[1,0,0,0]],[[290.000,450.000,10.000],[1.00000000,0.00000000,0.00000000,0.00000000]]];
		SuctionCup := [TRUE,[[-94.709,0.000,259.352],[0.00000000,0.00000000,0.00000000,1.00000000]],[1,[0,0,20],[1,0,0,0],0,0,0.005]];
		MoveAbsJ [[70.152800,32.938500,23.515600,0.000000,33.545900,70.152800],[9E+09,9E+09,9E+09,9E+09,9E+09,9E+09]],v1000,z1,SuctionCup \WObj:=In;
		MoveL [[-16.111,46.392,30.000],[0.00000000,1.00000000,0.00000000,-0.00000000],[0,2,-2,1],[9E+09,9E+09,9E+09,9E+09,9E+09,9E+09]],v1000,z1,SuctionCup \WObj:=In;
		! Attach to Suction Cup
		WaitTime 0.500;
		MoveL [[-16.087,46.472,70.960],[0.00000000,1.00000000,0.00000000,-0.00000000],[0,0,0,0],[9E+09,9E+09,9E+09,9E+09,9E+09,9E+09]],v1000,z1,SuctionCup \WObj:=In;
	ENDPROC

	PROC DropOut4()
		ConfJ \On;
		ConfL \Off;
		Out := [FALSE, TRUE, "", [[0,0,0],[1,0,0,0]],[[290.000,-450.000,10.000],[1.00000000,0.00000000,0.00000000,0.00000000]]];
		SuctionCup := [TRUE,[[-94.709,0.000,259.352],[0.00000000,0.00000000,0.00000000,1.00000000]],[1,[0,0,20],[1,0,0,0],0,0,0.005]];
		MoveAbsJ [[-66.056500,21.575200,36.080800,0.000000,32.344000,-66.056500],[9E+09,9E+09,9E+09,9E+09,9E+09,9E+09]],v1000,z1,SuctionCup \WObj:=Out;
		MoveL [[-16.111,46.392,45.000],[0.00000000,1.00000000,0.00000000,-0.00000000],[-1,0,-1,0],[9E+09,9E+09,9E+09,9E+09,9E+09,9E+09]],v1000,z1,SuctionCup \WObj:=Out;
		! Detach from Suction Cup
		WaitTime 0.500;
		MoveL [[-16.111,46.485,105.701],[0.00000000,1.00000000,0.00000000,-0.00000000],[-1,0,-1,0],[9E+09,9E+09,9E+09,9E+09,9E+09,9E+09]],v1000,z1,SuctionCup \WObj:=Out;
	ENDPROC

	PROC Main()
		ConfJ \On;
		ConfL \Off;
		! Program generated by VerticalBot Studio for ABB IRB 1200-5/0.9 on 25/10/2026 12:00:00
		! Using nominal kinematics.
		GoHome;
		PickIn1;
		GoHome;
		GoHome;
		DropStation;
		GoHome;
		Station1;
		GoHome;
		PickStation;
		GoHome;
		DropOut1;
		GoHome;
		PickIn2;
		GoHome;
		GoHome;
		DropStation;
		GoHome;
		Station1;
		GoHome;
		PickStation;
		GoHome;
		DropOut2;
		GoHome;
		PickIn3;
		GoHome;
		GoHome;
		DropStation;
		GoHome;
		Station1;
		GoHome;
		PickStation;
		GoHome;
		DropOut3;
		GoHome;
		PickIn4;
		GoHome;
		GoHome;
		DropStation;
		GoHome;
		Station1;
		GoHome;
		PickStation;
		GoHome;
		DropOut4;
		GoHome;
	ENDPROC

ENDMODULE
